(* Logix 5000 project; controller CIP_14485201 vendor 1 type 14 code 216 rev 38.11; software revision 38.01; part 2 of 12 *)

        [3].Setpoint[7] := 53.0, [3].Setpoint[8] := 63.0, [3].Setpoint[9] := 57.0, [3].Setpoint[10] := 43.0, [3].Setpoint[11] := 63.0, [3].Setpoint[13] := 85.0, [3].Setpoint[14] := 300.0, [3].Setpoint[15] := 900.0, [3].Setpoint[17] := 15.0, [3].Setpoint[18] := 14.0, [3].Setpoint[19] := 15.0, [3].Setpoint[20] := 45.0, [3].Setpoint[21] := 5.0, [3].Setpoint[22] := 15.0, [3].Setpoint[23] := 300.0, [3].Setpoint[25] := 10.0, [3].Setpoint[26] := 9.0, [3].Setpoint[27] := 10.0, [3].Setpoint[28] := 50.0, [3].Setpoint[29] := 3.0, [3].Setpoint[30] := 17.0, [3].Setpoint[31] := 300.0, [3].Setpoint[33] := 2.0, [3].Setpoint[34] := 900.0, [3].Setpoint[37] := 35.0, [3].Setpoint[41] := 5.0, [3].Setpoint[42] := 50.0, [3].Setpoint[43] := 5.0, [3].Setpoint[44] := 60.0, [3].Setpoint[45] := 50.0, [3].Setpoint[47] := 15.0, [3].Setpoint[49] := 180.0, [3].Setpoint[50] := 180.0, [3].Setpoint[52] := 30.0, [3].Setpoint[53] := 5.0, [3].Setpoint[54] := 5.0, [3].Setpoint[55] := 3.0, [3].Setpoint[57] := 300.0, [3].Name := 'RECIPE #3', [4].Setpoint[1] := 55.0, [4].Setpoint[2] := 65.0, [4].Setpoint[3] := 60.0, [4].Setpoint[4] := 45.0, [4].Setpoint[5] := 65.0, [4].Setpoint[7] := 53.0, [4].Setpoint[8] := 63.0, [4].Setpoint[9] := 57.0, [4].Setpoint[10] := 43.0, [4].Setpoint[11] := 63.0, [4].Setpoint[13] := 85.0, [4].Setpoint[14] := 300.0, [4].Setpoint[15] := 900.0, [4].Setpoint[17] := 15.0, [4].Setpoint[18] := 14.0, [4].Setpoint[19] := 15.0, [4].Setpoint[20] := 45.0, [4].Setpoint[21] := 5.0, [4].Setpoint[22] := 15.0, [4].Setpoint[23] := 300.0, [4].Setpoint[25] := 10.0,
        [4].Setpoint[26] := 9.0, [4].Setpoint[27] := 10.0, [4].Setpoint[28] := 50.0, [4].Setpoint[29] := 3.0, [4].Setpoint[30] := 17.0, [4].Setpoint[31] := 300.0, [4].Setpoint[33] := 2.0, [4].Setpoint[34] := 900.0, [4].Setpoint[37] := 35.0, [4].Setpoint[41] := 5.0, [4].Setpoint[42] := 50.0, [4].Setpoint[43] := 5.0, [4].Setpoint[44] := 60.0, [4].Setpoint[45] := 50.0, [4].Setpoint[47] := 15.0, [4].Setpoint[49] := 180.0, [4].Setpoint[50] := 180.0, [4].Setpoint[52] := 30.0, [4].Setpoint[53] := 5.0, [4].Setpoint[54] := 5.0, [4].Setpoint[55] := 3.0, [4].Setpoint[57] := 300.0, [4].Name := 'RECIPE #4', [5].Setpoint[1] := 55.0, [5].Setpoint[2] := 65.0, [5].Setpoint[3] := 60.0, [5].Setpoint[4] := 45.0, [5].Setpoint[5] := 65.0, [5].Setpoint[7] := 53.0, [5].Setpoint[8] := 63.0, [5].Setpoint[9] := 57.0, [5].Setpoint[10] := 43.0, [5].Setpoint[11] := 63.0, [5].Setpoint[13] := 85.0, [5].Setpoint[14] := 300.0, [5].Setpoint[15] := 900.0, [5].Setpoint[17] := 15.0, [5].Setpoint[18] := 14.0, [5].Setpoint[19] := 15.0, [5].Setpoint[20] := 45.0, [5].Setpoint[21] := 5.0, [5].Setpoint[22] := 15.0, [5].Setpoint[23] := 300.0, [5].Setpoint[25] := 10.0, [5].Setpoint[26] := 9.0, [5].Setpoint[27] := 10.0, [5].Setpoint[28] := 50.0, [5].Setpoint[29] := 3.0, [5].Setpoint[30] := 17.0, [5].Setpoint[31] := 300.0, [5].Setpoint[33] := 2.0, [5].Setpoint[34] := 900.0, [5].Setpoint[37] := 35.0, [5].Setpoint[41] := 5.0, [5].Setpoint[42] := 50.0, [5].Setpoint[43] := 5.0, [5].Setpoint[44] := 60.0, [5].Setpoint[45] := 50.0, [5].Setpoint[47] := 15.0, [5].Setpoint[49] := 180.0,
        [5].Setpoint[50] := 180.0, [5].Setpoint[52] := 30.0, [5].Setpoint[53] := 5.0, [5].Setpoint[54] := 5.0, [5].Setpoint[55] := 3.0, [5].Setpoint[57] := 300.0, [5].Name := 'RECIPE #5', [6].Setpoint[1] := 55.0, [6].Setpoint[2] := 65.0, [6].Setpoint[3] := 60.0, [6].Setpoint[4] := 45.0, [6].Setpoint[5] := 65.0, [6].Setpoint[7] := 53.0, [6].Setpoint[8] := 63.0, [6].Setpoint[9] := 57.0, [6].Setpoint[10] := 43.0, [6].Setpoint[11] := 63.0, [6].Setpoint[13] := 85.0, [6].Setpoint[14] := 300.0, [6].Setpoint[15] := 900.0, [6].Setpoint[17] := 15.0, [6].Setpoint[18] := 14.0, [6].Setpoint[19] := 15.0, [6].Setpoint[20] := 45.0, [6].Setpoint[21] := 5.0, [6].Setpoint[22] := 15.0, [6].Setpoint[23] := 300.0, [6].Setpoint[25] := 10.0, [6].Setpoint[26] := 9.0, [6].Setpoint[27] := 10.0, [6].Setpoint[28] := 50.0, [6].Setpoint[29] := 3.0, [6].Setpoint[30] := 17.0, [6].Setpoint[31] := 300.0, [6].Setpoint[33] := 2.0, [6].Setpoint[34] := 900.0, [6].Setpoint[37] := 35.0, [6].Setpoint[41] := 5.0, [6].Setpoint[42] := 50.0, [6].Setpoint[43] := 5.0, [6].Setpoint[44] := 60.0, [6].Setpoint[45] := 50.0, [6].Setpoint[47] := 15.0, [6].Setpoint[49] := 180.0, [6].Setpoint[50] := 180.0, [6].Setpoint[52] := 30.0, [6].Setpoint[53] := 5.0, [6].Setpoint[54] := 5.0, [6].Setpoint[55] := 3.0, [6].Setpoint[57] := 300.0, [6].Name := 'RECIPE #6', [7].Setpoint[1] := 55.0, [7].Setpoint[2] := 65.0, [7].Setpoint[3] := 60.0, [7].Setpoint[4] := 45.0, [7].Setpoint[5] := 65.0, [7].Setpoint[7] := 53.0, [7].Setpoint[8] := 63.0, [7].Setpoint[9] := 57.0, [7].Setpoint[10] := 43.0,
        [7].Setpoint[11] := 63.0, [7].Setpoint[13] := 85.0, [7].Setpoint[14] := 300.0, [7].Setpoint[15] := 900.0, [7].Setpoint[17] := 15.0, [7].Setpoint[18] := 14.0, [7].Setpoint[19] := 15.0, [7].Setpoint[20] := 45.0, [7].Setpoint[21] := 5.0, [7].Setpoint[22] := 15.0, [7].Setpoint[23] := 300.0, [7].Setpoint[25] := 10.0, [7].Setpoint[26] := 9.0, [7].Setpoint[27] := 10.0, [7].Setpoint[28] := 50.0, [7].Setpoint[29] := 3.0, [7].Setpoint[30] := 17.0, [7].Setpoint[31] := 300.0, [7].Setpoint[33] := 2.0, [7].Setpoint[34] := 900.0, [7].Setpoint[37] := 35.0, [7].Setpoint[41] := 5.0, [7].Setpoint[42] := 50.0, [7].Setpoint[43] := 5.0, [7].Setpoint[44] := 60.0, [7].Setpoint[45] := 50.0, [7].Setpoint[47] := 15.0, [7].Setpoint[49] := 180.0, [7].Setpoint[50] := 180.0, [7].Setpoint[52] := 30.0, [7].Setpoint[53] := 5.0, [7].Setpoint[54] := 5.0, [7].Setpoint[55] := 3.0, [7].Setpoint[57] := 300.0, [7].Name := 'RECIPE #7', [8].Setpoint[1] := 55.0, [8].Setpoint[2] := 65.0, [8].Setpoint[3] := 60.0, [8].Setpoint[4] := 45.0, [8].Setpoint[5] := 65.0, [8].Setpoint[7] := 53.0, [8].Setpoint[8] := 63.0, [8].Setpoint[9] := 57.0, [8].Setpoint[10] := 43.0, [8].Setpoint[11] := 63.0, [8].Setpoint[13] := 85.0, [8].Setpoint[14] := 300.0, [8].Setpoint[15] := 900.0, [8].Setpoint[17] := 15.0, [8].Setpoint[18] := 14.0, [8].Setpoint[19] := 15.0, [8].Setpoint[20] := 45.0, [8].Setpoint[21] := 5.0, [8].Setpoint[22] := 15.0, [8].Setpoint[23] := 300.0, [8].Setpoint[25] := 10.0, [8].Setpoint[26] := 9.0, [8].Setpoint[27] := 10.0, [8].Setpoint[28] := 50.0, [8].Setpoint[29] := 3.0,
        [8].Setpoint[30] := 17.0, [8].Setpoint[31] := 300.0, [8].Setpoint[33] := 2.0, [8].Setpoint[34] := 900.0, [8].Setpoint[37] := 35.0, [8].Setpoint[41] := 5.0, [8].Setpoint[42] := 50.0, [8].Setpoint[43] := 5.0, [8].Setpoint[44] := 60.0, [8].Setpoint[45] := 50.0, [8].Setpoint[47] := 15.0, [8].Setpoint[49] := 180.0, [8].Setpoint[50] := 180.0, [8].Setpoint[52] := 30.0, [8].Setpoint[53] := 5.0, [8].Setpoint[54] := 5.0, [8].Setpoint[55] := 3.0, [8].Setpoint[57] := 300.0, [8].Name := 'RECIPE #8', [9].Setpoint[1] := 55.0, [9].Setpoint[2] := 65.0, [9].Setpoint[3] := 60.0, [9].Setpoint[4] := 45.0, [9].Setpoint[5] := 65.0, [9].Setpoint[7] := 53.0, [9].Setpoint[8] := 63.0, [9].Setpoint[9] := 57.0, [9].Setpoint[10] := 43.0, [9].Setpoint[11] := 63.0, [9].Setpoint[13] := 85.0, [9].Setpoint[14] := 300.0, [9].Setpoint[15] := 900.0, [9].Setpoint[17] := 15.0, [9].Setpoint[18] := 14.0, [9].Setpoint[19] := 15.0, [9].Setpoint[20] := 45.0, [9].Setpoint[21] := 5.0, [9].Setpoint[22] := 15.0, [9].Setpoint[23] := 300.0, [9].Setpoint[25] := 10.0, [9].Setpoint[26] := 9.0, [9].Setpoint[27] := 10.0, [9].Setpoint[28] := 50.0, [9].Setpoint[29] := 3.0, [9].Setpoint[30] := 17.0, [9].Setpoint[31] := 300.0, [9].Setpoint[33] := 2.0, [9].Setpoint[34] := 900.0, [9].Setpoint[37] := 35.0, [9].Setpoint[41] := 5.0, [9].Setpoint[42] := 50.0, [9].Setpoint[43] := 5.0, [9].Setpoint[44] := 60.0, [9].Setpoint[45] := 50.0, [9].Setpoint[47] := 15.0, [9].Setpoint[49] := 180.0, [9].Setpoint[50] := 180.0, [9].Setpoint[52] := 30.0, [9].Setpoint[53] := 5.0, [9].Setpoint[54] := 5.0,
        [9].Setpoint[55] := 3.0, [9].Setpoint[57] := 300.0, [9].Name := 'RECIPE #9', [10].Setpoint[1] := 55.0, [10].Setpoint[2] := 65.0, [10].Setpoint[3] := 60.0, [10].Setpoint[4] := 45.0, [10].Setpoint[5] := 65.0, [10].Setpoint[7] := 53.0, [10].Setpoint[8] := 63.0, [10].Setpoint[9] := 57.0, [10].Setpoint[10] := 43.0, [10].Setpoint[11] := 63.0, [10].Setpoint[13] := 85.0, [10].Setpoint[14] := 300.0, [10].Setpoint[15] := 900.0, [10].Setpoint[17] := 15.0, [10].Setpoint[18] := 14.0, [10].Setpoint[19] := 15.0, [10].Setpoint[20] := 45.0, [10].Setpoint[21] := 5.0, [10].Setpoint[22] := 15.0, [10].Setpoint[23] := 300.0, [10].Setpoint[25] := 10.0, [10].Setpoint[26] := 9.0, [10].Setpoint[27] := 10.0, [10].Setpoint[28] := 50.0, [10].Setpoint[29] := 3.0, [10].Setpoint[30] := 17.0, [10].Setpoint[31] := 300.0, [10].Setpoint[33] := 2.0, [10].Setpoint[34] := 900.0, [10].Setpoint[37] := 35.0, [10].Setpoint[41] := 5.0, [10].Setpoint[42] := 50.0, [10].Setpoint[43] := 5.0, [10].Setpoint[44] := 60.0, [10].Setpoint[45] := 50.0, [10].Setpoint[47] := 15.0, [10].Setpoint[49] := 180.0, [10].Setpoint[50] := 180.0, [10].Setpoint[52] := 30.0, [10].Setpoint[53] := 5.0, [10].Setpoint[54] := 5.0, [10].Setpoint[55] := 3.0, [10].Setpoint[57] := 300.0, [10].Name := 'RECIPE #10', [11].Setpoint[1] := 55.0, [11].Setpoint[2] := 65.0, [11].Setpoint[3] := 60.0, [11].Setpoint[4] := 45.0, [11].Setpoint[5] := 65.0, [11].Setpoint[7] := 53.0, [11].Setpoint[8] := 63.0, [11].Setpoint[9] := 57.0, [11].Setpoint[10] := 43.0, [11].Setpoint[11] := 63.0, [11].Setpoint[13] := 85.0, [11].Setpoint[14] := 300.0, [11].Setpoint[15] := 900.0,
        [11].Setpoint[17] := 15.0, [11].Setpoint[18] := 14.0, [11].Setpoint[19] := 15.0, [11].Setpoint[20] := 45.0, [11].Setpoint[21] := 5.0, [11].Setpoint[22] := 15.0, [11].Setpoint[23] := 300.0, [11].Setpoint[25] := 10.0, [11].Setpoint[26] := 9.0, [11].Setpoint[27] := 10.0, [11].Setpoint[28] := 50.0, [11].Setpoint[29] := 3.0, [11].Setpoint[30] := 17.0, [11].Setpoint[31] := 300.0, [11].Setpoint[33] := 2.0, [11].Setpoint[34] := 900.0, [11].Setpoint[37] := 35.0, [11].Setpoint[41] := 5.0, [11].Setpoint[42] := 50.0, [11].Setpoint[43] := 5.0, [11].Setpoint[44] := 60.0, [11].Setpoint[45] := 50.0, [11].Setpoint[47] := 15.0, [11].Setpoint[49] := 180.0, [11].Setpoint[50] := 180.0, [11].Setpoint[52] := 30.0, [11].Setpoint[53] := 5.0, [11].Setpoint[54] := 5.0, [11].Setpoint[55] := 3.0, [11].Setpoint[57] := 300.0, [11].Name := 'RECIPE #11', [12].Setpoint[1] := 55.0, [12].Setpoint[2] := 65.0, [12].Setpoint[3] := 60.0, [12].Setpoint[4] := 45.0, [12].Setpoint[5] := 65.0, [12].Setpoint[7] := 53.0, [12].Setpoint[8] := 63.0, [12].Setpoint[9] := 57.0, [12].Setpoint[10] := 43.0, [12].Setpoint[11] := 63.0, [12].Setpoint[13] := 85.0, [12].Setpoint[14] := 300.0, [12].Setpoint[15] := 900.0, [12].Setpoint[17] := 15.0, [12].Setpoint[18] := 14.0, [12].Setpoint[19] := 15.0, [12].Setpoint[20] := 45.0, [12].Setpoint[21] := 5.0, [12].Setpoint[22] := 15.0, [12].Setpoint[23] := 300.0, [12].Setpoint[25] := 10.0, [12].Setpoint[26] := 9.0, [12].Setpoint[27] := 10.0, [12].Setpoint[28] := 50.0, [12].Setpoint[29] := 3.0, [12].Setpoint[30] := 17.0, [12].Setpoint[31] := 300.0, [12].Setpoint[33] := 2.0, [12].Setpoint[34] := 900.0,
        [12].Setpoint[37] := 35.0, [12].Setpoint[41] := 5.0, [12].Setpoint[42] := 50.0, [12].Setpoint[43] := 5.0, [12].Setpoint[44] := 60.0, [12].Setpoint[45] := 50.0, [12].Setpoint[47] := 15.0, [12].Setpoint[49] := 180.0, [12].Setpoint[50] := 180.0, [12].Setpoint[52] := 30.0, [12].Setpoint[53] := 5.0, [12].Setpoint[54] := 5.0, [12].Setpoint[55] := 3.0, [12].Setpoint[57] := 300.0, [12].Name := 'RECIPE #12', [13].Setpoint[1] := 55.0, [13].Setpoint[2] := 65.0, [13].Setpoint[3] := 60.0, [13].Setpoint[4] := 45.0, [13].Setpoint[5] := 65.0, [13].Setpoint[7] := 53.0, [13].Setpoint[8] := 63.0, [13].Setpoint[9] := 57.0, [13].Setpoint[10] := 43.0, [13].Setpoint[11] := 63.0, [13].Setpoint[13] := 85.0, [13].Setpoint[14] := 300.0, [13].Setpoint[15] := 900.0, [13].Setpoint[17] := 15.0, [13].Setpoint[18] := 14.0, [13].Setpoint[19] := 15.0, [13].Setpoint[20] := 45.0, [13].Setpoint[21] := 5.0, [13].Setpoint[22] := 15.0, [13].Setpoint[23] := 300.0, [13].Setpoint[25] := 10.0, [13].Setpoint[26] := 9.0, [13].Setpoint[27] := 10.0, [13].Setpoint[28] := 50.0, [13].Setpoint[29] := 3.0, [13].Setpoint[30] := 17.0, [13].Setpoint[31] := 300.0, [13].Setpoint[33] := 2.0, [13].Setpoint[34] := 900.0, [13].Setpoint[37] := 35.0, [13].Setpoint[41] := 5.0, [13].Setpoint[42] := 50.0, [13].Setpoint[43] := 5.0, [13].Setpoint[44] := 60.0, [13].Setpoint[45] := 50.0, [13].Setpoint[47] := 15.0, [13].Setpoint[49] := 180.0, [13].Setpoint[50] := 180.0, [13].Setpoint[52] := 30.0, [13].Setpoint[53] := 5.0, [13].Setpoint[54] := 5.0, [13].Setpoint[55] := 3.0, [13].Setpoint[57] := 300.0, [13].Name := 'RECIPE #13', [14].Setpoint[1] := 55.0,
        [14].Setpoint[2] := 65.0, [14].Setpoint[3] := 60.0, [14].Setpoint[4] := 45.0, [14].Setpoint[5] := 65.0, [14].Setpoint[7] := 53.0, [14].Setpoint[8] := 63.0, [14].Setpoint[9] := 57.0, [14].Setpoint[10] := 43.0, [14].Setpoint[11] := 63.0, [14].Setpoint[13] := 85.0, [14].Setpoint[14] := 300.0, [14].Setpoint[15] := 900.0, [14].Setpoint[17] := 15.0, [14].Setpoint[18] := 14.0, [14].Setpoint[19] := 15.0, [14].Setpoint[20] := 45.0, [14].Setpoint[21] := 5.0, [14].Setpoint[22] := 15.0, [14].Setpoint[23] := 300.0, [14].Setpoint[25] := 10.0, [14].Setpoint[26] := 9.0, [14].Setpoint[27] := 10.0, [14].Setpoint[28] := 50.0, [14].Setpoint[29] := 3.0, [14].Setpoint[30] := 17.0, [14].Setpoint[31] := 300.0, [14].Setpoint[33] := 2.0, [14].Setpoint[34] := 900.0, [14].Setpoint[37] := 35.0, [14].Setpoint[41] := 5.0, [14].Setpoint[42] := 50.0, [14].Setpoint[43] := 5.0, [14].Setpoint[44] := 60.0, [14].Setpoint[45] := 50.0, [14].Setpoint[47] := 15.0, [14].Setpoint[49] := 180.0, [14].Setpoint[50] := 180.0, [14].Setpoint[52] := 30.0, [14].Setpoint[53] := 5.0, [14].Setpoint[54] := 5.0, [14].Setpoint[55] := 3.0, [14].Setpoint[57] := 300.0, [14].Name := 'RECIPE #14', [15].Setpoint[1] := 55.0, [15].Setpoint[2] := 65.0, [15].Setpoint[3] := 60.0, [15].Setpoint[4] := 45.0, [15].Setpoint[5] := 65.0, [15].Setpoint[7] := 53.0, [15].Setpoint[8] := 63.0, [15].Setpoint[9] := 57.0, [15].Setpoint[10] := 43.0, [15].Setpoint[11] := 63.0, [15].Setpoint[13] := 85.0, [15].Setpoint[14] := 300.0, [15].Setpoint[15] := 900.0, [15].Setpoint[17] := 15.0, [15].Setpoint[18] := 14.0, [15].Setpoint[19] := 15.0, [15].Setpoint[20] := 45.0,
        [15].Setpoint[21] := 5.0, [15].Setpoint[22] := 15.0, [15].Setpoint[23] := 300.0, [15].Setpoint[25] := 10.0, [15].Setpoint[26] := 9.0, [15].Setpoint[27] := 10.0, [15].Setpoint[28] := 50.0, [15].Setpoint[29] := 3.0, [15].Setpoint[30] := 17.0, [15].Setpoint[31] := 300.0, [15].Setpoint[33] := 2.0, [15].Setpoint[34] := 900.0, [15].Setpoint[37] := 35.0, [15].Setpoint[41] := 5.0, [15].Setpoint[42] := 50.0, [15].Setpoint[43] := 5.0, [15].Setpoint[44] := 60.0, [15].Setpoint[45] := 50.0, [15].Setpoint[47] := 15.0, [15].Setpoint[49] := 180.0, [15].Setpoint[50] := 180.0, [15].Setpoint[52] := 30.0, [15].Setpoint[53] := 5.0, [15].Setpoint[54] := 5.0, [15].Setpoint[55] := 3.0, [15].Setpoint[57] := 300.0, [15].Name := 'RECIPE #15', [16].Setpoint[1] := 55.0, [16].Setpoint[2] := 65.0, [16].Setpoint[3] := 60.0, [16].Setpoint[4] := 45.0, [16].Setpoint[5] := 65.0, [16].Setpoint[7] := 53.0, [16].Setpoint[8] := 63.0, [16].Setpoint[9] := 57.0, [16].Setpoint[10] := 43.0, [16].Setpoint[11] := 63.0, [16].Setpoint[13] := 85.0, [16].Setpoint[14] := 300.0, [16].Setpoint[15] := 900.0, [16].Setpoint[17] := 15.0, [16].Setpoint[18] := 14.0, [16].Setpoint[19] := 15.0, [16].Setpoint[20] := 45.0, [16].Setpoint[21] := 5.0, [16].Setpoint[22] := 15.0, [16].Setpoint[23] := 300.0, [16].Setpoint[25] := 10.0, [16].Setpoint[26] := 9.0, [16].Setpoint[27] := 10.0, [16].Setpoint[28] := 50.0, [16].Setpoint[29] := 3.0, [16].Setpoint[30] := 17.0, [16].Setpoint[31] := 300.0, [16].Setpoint[33] := 2.0, [16].Setpoint[34] := 900.0, [16].Setpoint[37] := 35.0, [16].Setpoint[41] := 5.0, [16].Setpoint[42] := 50.0, [16].Setpoint[43] := 5.0,
        [16].Setpoint[44] := 60.0, [16].Setpoint[45] := 50.0, [16].Setpoint[47] := 15.0, [16].Setpoint[49] := 180.0, [16].Setpoint[50] := 180.0, [16].Setpoint[52] := 30.0, [16].Setpoint[53] := 5.0, [16].Setpoint[54] := 5.0, [16].Setpoint[55] := 3.0, [16].Setpoint[57] := 300.0, [16].Name := 'RECIPE #16', [17].Setpoint[1] := 55.0, [17].Setpoint[2] := 65.0, [17].Setpoint[3] := 60.0, [17].Setpoint[4] := 45.0, [17].Setpoint[5] := 65.0, [17].Setpoint[7] := 53.0, [17].Setpoint[8] := 63.0, [17].Setpoint[9] := 57.0, [17].Setpoint[10] := 43.0, [17].Setpoint[11] := 63.0, [17].Setpoint[13] := 85.0, [17].Setpoint[14] := 300.0, [17].Setpoint[15] := 900.0, [17].Setpoint[17] := 15.0, [17].Setpoint[18] := 14.0, [17].Setpoint[19] := 15.0, [17].Setpoint[20] := 45.0, [17].Setpoint[21] := 5.0, [17].Setpoint[22] := 15.0, [17].Setpoint[23] := 300.0, [17].Setpoint[25] := 10.0, [17].Setpoint[26] := 9.0, [17].Setpoint[27] := 10.0, [17].Setpoint[28] := 50.0, [17].Setpoint[29] := 3.0, [17].Setpoint[30] := 17.0, [17].Setpoint[31] := 300.0, [17].Setpoint[33] := 2.0, [17].Setpoint[34] := 900.0, [17].Setpoint[37] := 35.0, [17].Setpoint[41] := 5.0, [17].Setpoint[42] := 50.0, [17].Setpoint[43] := 5.0, [17].Setpoint[44] := 60.0, [17].Setpoint[45] := 50.0, [17].Setpoint[47] := 15.0, [17].Setpoint[49] := 180.0, [17].Setpoint[50] := 180.0, [17].Setpoint[52] := 30.0, [17].Setpoint[53] := 5.0, [17].Setpoint[54] := 5.0, [17].Setpoint[55] := 3.0, [17].Setpoint[57] := 300.0, [17].Name := 'RECIPE #17', [18].Setpoint[1] := 55.0, [18].Setpoint[2] := 65.0, [18].Setpoint[3] := 60.0, [18].Setpoint[4] := 45.0, [18].Setpoint[5] := 65.0,
        [18].Setpoint[7] := 53.0, [18].Setpoint[8] := 63.0, [18].Setpoint[9] := 57.0, [18].Setpoint[10] := 43.0, [18].Setpoint[11] := 63.0, [18].Setpoint[13] := 85.0, [18].Setpoint[14] := 300.0, [18].Setpoint[15] := 900.0, [18].Setpoint[17] := 15.0, [18].Setpoint[18] := 14.0, [18].Setpoint[19] := 15.0, [18].Setpoint[20] := 45.0, [18].Setpoint[21] := 5.0, [18].Setpoint[22] := 15.0, [18].Setpoint[23] := 300.0, [18].Setpoint[25] := 10.0, [18].Setpoint[26] := 9.0, [18].Setpoint[27] := 10.0, [18].Setpoint[28] := 50.0, [18].Setpoint[29] := 3.0, [18].Setpoint[30] := 17.0, [18].Setpoint[31] := 300.0, [18].Setpoint[33] := 2.0, [18].Setpoint[34] := 900.0, [18].Setpoint[37] := 35.0, [18].Setpoint[41] := 5.0, [18].Setpoint[42] := 50.0, [18].Setpoint[43] := 5.0, [18].Setpoint[44] := 60.0, [18].Setpoint[45] := 50.0, [18].Setpoint[47] := 15.0, [18].Setpoint[49] := 180.0, [18].Setpoint[50] := 180.0, [18].Setpoint[52] := 30.0, [18].Setpoint[53] := 5.0, [18].Setpoint[54] := 5.0, [18].Setpoint[55] := 3.0, [18].Setpoint[57] := 300.0, [18].Name := 'RECIPE #18', [19].Setpoint[1] := 55.0, [19].Setpoint[2] := 65.0, [19].Setpoint[3] := 60.0, [19].Setpoint[4] := 45.0, [19].Setpoint[5] := 65.0, [19].Setpoint[7] := 53.0, [19].Setpoint[8] := 63.0, [19].Setpoint[9] := 57.0, [19].Setpoint[10] := 43.0, [19].Setpoint[11] := 63.0, [19].Setpoint[13] := 85.0, [19].Setpoint[14] := 300.0, [19].Setpoint[15] := 900.0, [19].Setpoint[17] := 15.0, [19].Setpoint[18] := 14.0, [19].Setpoint[19] := 15.0, [19].Setpoint[20] := 45.0, [19].Setpoint[21] := 5.0, [19].Setpoint[22] := 15.0, [19].Setpoint[23] := 300.0, [19].Setpoint[25] := 10.0,
        [19].Setpoint[26] := 9.0, [19].Setpoint[27] := 10.0, [19].Setpoint[28] := 50.0, [19].Setpoint[29] := 3.0, [19].Setpoint[30] := 17.0, [19].Setpoint[31] := 300.0, [19].Setpoint[33] := 2.0, [19].Setpoint[34] := 900.0, [19].Setpoint[37] := 35.0, [19].Setpoint[41] := 5.0, [19].Setpoint[42] := 50.0, [19].Setpoint[43] := 5.0, [19].Setpoint[44] := 60.0, [19].Setpoint[45] := 50.0, [19].Setpoint[47] := 15.0, [19].Setpoint[49] := 180.0, [19].Setpoint[50] := 180.0, [19].Setpoint[52] := 30.0, [19].Setpoint[53] := 5.0, [19].Setpoint[54] := 5.0, [19].Setpoint[55] := 3.0, [19].Setpoint[57] := 300.0, [19].Name := 'RECIPE #19', [20].Setpoint[1] := 55.0, [20].Setpoint[2] := 65.0, [20].Setpoint[3] := 60.0, [20].Setpoint[4] := 45.0, [20].Setpoint[5] := 65.0, [20].Setpoint[7] := 53.0, [20].Setpoint[8] := 63.0, [20].Setpoint[9] := 57.0, [20].Setpoint[10] := 43.0, [20].Setpoint[11] := 63.0, [20].Setpoint[13] := 85.0, [20].Setpoint[14] := 300.0, [20].Setpoint[15] := 900.0, [20].Setpoint[17] := 15.0, [20].Setpoint[18] := 14.0, [20].Setpoint[19] := 15.0, [20].Setpoint[20] := 45.0, [20].Setpoint[21] := 5.0, [20].Setpoint[22] := 15.0, [20].Setpoint[23] := 300.0, [20].Setpoint[25] := 10.0, [20].Setpoint[26] := 9.0, [20].Setpoint[27] := 10.0, [20].Setpoint[28] := 50.0, [20].Setpoint[29] := 3.0, [20].Setpoint[30] := 17.0, [20].Setpoint[31] := 300.0, [20].Setpoint[33] := 2.0, [20].Setpoint[34] := 900.0, [20].Setpoint[37] := 35.0, [20].Setpoint[41] := 5.0, [20].Setpoint[42] := 50.0, [20].Setpoint[43] := 5.0, [20].Setpoint[44] := 60.0, [20].Setpoint[45] := 50.0, [20].Setpoint[47] := 15.0, [20].Setpoint[49] := 180.0,
        [20].Setpoint[50] := 180.0, [20].Setpoint[52] := 30.0, [20].Setpoint[53] := 5.0, [20].Setpoint[54] := 5.0, [20].Setpoint[55] := 3.0, [20].Setpoint[57] := 300.0, [20].Name := 'RECIPE #20', [21].Setpoint[1] := 55.0, [21].Setpoint[2] := 65.0, [21].Setpoint[3] := 60.0, [21].Setpoint[4] := 45.0, [21].Setpoint[5] := 65.0, [21].Setpoint[7] := 53.0, [21].Setpoint[8] := 63.0, [21].Setpoint[9] := 57.0, [21].Setpoint[10] := 43.0, [21].Setpoint[11] := 63.0, [21].Setpoint[13] := 85.0, [21].Setpoint[14] := 300.0, [21].Setpoint[15] := 900.0, [21].Setpoint[17] := 15.0, [21].Setpoint[18] := 14.0, [21].Setpoint[19] := 15.0, [21].Setpoint[20] := 45.0, [21].Setpoint[21] := 5.0, [21].Setpoint[22] := 15.0, [21].Setpoint[23] := 300.0, [21].Setpoint[25] := 10.0, [21].Setpoint[26] := 9.0, [21].Setpoint[27] := 10.0, [21].Setpoint[28] := 50.0, [21].Setpoint[29] := 3.0, [21].Setpoint[30] := 17.0, [21].Setpoint[31] := 300.0, [21].Setpoint[33] := 2.0, [21].Setpoint[34] := 900.0, [21].Setpoint[37] := 35.0, [21].Setpoint[41] := 5.0, [21].Setpoint[42] := 50.0, [21].Setpoint[43] := 5.0, [21].Setpoint[44] := 60.0, [21].Setpoint[45] := 50.0, [21].Setpoint[47] := 15.0, [21].Setpoint[49] := 180.0, [21].Setpoint[50] := 180.0, [21].Setpoint[52] := 30.0, [21].Setpoint[53] := 5.0, [21].Setpoint[54] := 5.0, [21].Setpoint[55] := 3.0, [21].Setpoint[57] := 300.0, [21].Name := 'RECIPE #21', [22].Setpoint[1] := 55.0, [22].Setpoint[2] := 65.0, [22].Setpoint[3] := 60.0, [22].Setpoint[4] := 45.0, [22].Setpoint[5] := 65.0, [22].Setpoint[7] := 53.0, [22].Setpoint[8] := 63.0, [22].Setpoint[9] := 57.0, [22].Setpoint[10] := 43.0,
        [22].Setpoint[11] := 63.0, [22].Setpoint[13] := 85.0, [22].Setpoint[14] := 300.0, [22].Setpoint[15] := 900.0, [22].Setpoint[17] := 15.0, [22].Setpoint[18] := 14.0, [22].Setpoint[19] := 15.0, [22].Setpoint[20] := 45.0, [22].Setpoint[21] := 5.0, [22].Setpoint[22] := 15.0, [22].Setpoint[23] := 300.0, [22].Setpoint[25] := 10.0, [22].Setpoint[26] := 9.0, [22].Setpoint[27] := 10.0, [22].Setpoint[28] := 50.0, [22].Setpoint[29] := 3.0, [22].Setpoint[30] := 17.0, [22].Setpoint[31] := 300.0, [22].Setpoint[33] := 2.0, [22].Setpoint[34] := 900.0, [22].Setpoint[37] := 35.0, [22].Setpoint[41] := 5.0, [22].Setpoint[42] := 50.0, [22].Setpoint[43] := 5.0, [22].Setpoint[44] := 60.0, [22].Setpoint[45] := 50.0, [22].Setpoint[47] := 15.0, [22].Setpoint[49] := 180.0, [22].Setpoint[50] := 180.0, [22].Setpoint[52] := 30.0, [22].Setpoint[53] := 5.0, [22].Setpoint[54] := 5.0, [22].Setpoint[55] := 3.0, [22].Setpoint[57] := 300.0, [22].Name := 'RECIPE #22', [23].Setpoint[1] := 55.0, [23].Setpoint[2] := 65.0, [23].Setpoint[3] := 60.0, [23].Setpoint[4] := 45.0, [23].Setpoint[5] := 65.0, [23].Setpoint[7] := 53.0, [23].Setpoint[8] := 63.0, [23].Setpoint[9] := 57.0, [23].Setpoint[10] := 43.0, [23].Setpoint[11] := 63.0, [23].Setpoint[13] := 85.0, [23].Setpoint[14] := 300.0, [23].Setpoint[15] := 900.0, [23].Setpoint[17] := 15.0, [23].Setpoint[18] := 14.0, [23].Setpoint[19] := 15.0, [23].Setpoint[20] := 45.0, [23].Setpoint[21] := 5.0, [23].Setpoint[22] := 15.0, [23].Setpoint[23] := 300.0, [23].Setpoint[25] := 10.0, [23].Setpoint[26] := 9.0, [23].Setpoint[27] := 10.0, [23].Setpoint[28] := 50.0, [23].Setpoint[29] := 3.0,
        [23].Setpoint[30] := 17.0, [23].Setpoint[31] := 300.0, [23].Setpoint[33] := 2.0, [23].Setpoint[34] := 900.0, [23].Setpoint[37] := 35.0, [23].Setpoint[41] := 5.0, [23].Setpoint[42] := 50.0, [23].Setpoint[43] := 5.0, [23].Setpoint[44] := 60.0, [23].Setpoint[45] := 50.0, [23].Setpoint[47] := 15.0, [23].Setpoint[49] := 180.0, [23].Setpoint[50] := 180.0, [23].Setpoint[52] := 30.0, [23].Setpoint[53] := 5.0, [23].Setpoint[54] := 5.0, [23].Setpoint[55] := 3.0, [23].Setpoint[57] := 300.0, [23].Name := 'RECIPE #23', [24].OpCode[88] := 2, [24].Setpoint[1] := 55.0, [24].Setpoint[2] := 65.0, [24].Setpoint[3] := 60.0, [24].Setpoint[4] := 45.0, [24].Setpoint[5] := 65.0, [24].Setpoint[7] := 53.0, [24].Setpoint[8] := 63.0, [24].Setpoint[9] := 57.0, [24].Setpoint[10] := 43.0, [24].Setpoint[11] := 63.0, [24].Setpoint[13] := 85.0, [24].Setpoint[14] := 300.0, [24].Setpoint[15] := 900.0, [24].Setpoint[17] := 15.0, [24].Setpoint[18] := 14.0, [24].Setpoint[19] := 15.0, [24].Setpoint[20] := 45.0, [24].Setpoint[21] := 5.0, [24].Setpoint[22] := 15.0, [24].Setpoint[23] := 300.0, [24].Setpoint[25] := 10.0, [24].Setpoint[26] := 9.0, [24].Setpoint[27] := 10.0, [24].Setpoint[28] := 50.0, [24].Setpoint[29] := 3.0, [24].Setpoint[30] := 17.0, [24].Setpoint[31] := 300.0, [24].Setpoint[33] := 2.0, [24].Setpoint[34] := 900.0, [24].Setpoint[37] := 35.0, [24].Setpoint[41] := 5.0, [24].Setpoint[42] := 50.0, [24].Setpoint[43] := 5.0, [24].Setpoint[44] := 60.0, [24].Setpoint[45] := 50.0, [24].Setpoint[47] := 15.0, [24].Setpoint[49] := 180.0, [24].Setpoint[50] := 180.0, [24].Setpoint[52] := 30.0, [24].Setpoint[53] := 5.0,
        [24].Setpoint[54] := 5.0, [24].Setpoint[55] := 3.0, [24].Setpoint[57] := 300.0, [24].Name := 'RECIPE #24', [25].Setpoint[1] := 55.0, [25].Setpoint[2] := 65.0, [25].Setpoint[3] := 60.0, [25].Setpoint[4] := 45.0, [25].Setpoint[5] := 65.0, [25].Setpoint[7] := 53.0, [25].Setpoint[8] := 63.0, [25].Setpoint[9] := 57.0, [25].Setpoint[10] := 43.0, [25].Setpoint[11] := 63.0, [25].Setpoint[13] := 85.0, [25].Setpoint[14] := 300.0, [25].Setpoint[15] := 900.0, [25].Setpoint[17] := 15.0, [25].Setpoint[18] := 14.0, [25].Setpoint[19] := 15.0, [25].Setpoint[20] := 45.0, [25].Setpoint[21] := 5.0, [25].Setpoint[22] := 15.0, [25].Setpoint[23] := 300.0, [25].Setpoint[25] := 10.0, [25].Setpoint[26] := 9.0, [25].Setpoint[27] := 10.0, [25].Setpoint[28] := 50.0, [25].Setpoint[29] := 3.0, [25].Setpoint[30] := 17.0, [25].Setpoint[31] := 300.0, [25].Setpoint[33] := 2.0, [25].Setpoint[34] := 900.0, [25].Setpoint[37] := 35.0, [25].Setpoint[41] := 5.0, [25].Setpoint[42] := 50.0, [25].Setpoint[43] := 5.0, [25].Setpoint[44] := 60.0, [25].Setpoint[45] := 50.0, [25].Setpoint[47] := 15.0, [25].Setpoint[49] := 180.0, [25].Setpoint[50] := 180.0, [25].Setpoint[52] := 30.0, [25].Setpoint[53] := 5.0, [25].Setpoint[54] := 5.0, [25].Setpoint[55] := 3.0, [25].Setpoint[57] := 300.0, [25].Name := 'RECIPE #25', [26].Setpoint[1] := 55.0, [26].Setpoint[2] := 65.0, [26].Setpoint[3] := 60.0, [26].Setpoint[4] := 45.0, [26].Setpoint[5] := 65.0, [26].Setpoint[7] := 53.0, [26].Setpoint[8] := 63.0, [26].Setpoint[9] := 57.0, [26].Setpoint[10] := 43.0, [26].Setpoint[11] := 63.0, [26].Setpoint[13] := 85.0, [26].Setpoint[14] := 300.0,
        [26].Setpoint[15] := 900.0, [26].Setpoint[17] := 15.0, [26].Setpoint[18] := 14.0, [26].Setpoint[19] := 15.0, [26].Setpoint[20] := 45.0, [26].Setpoint[21] := 5.0, [26].Setpoint[22] := 15.0, [26].Setpoint[23] := 300.0, [26].Setpoint[25] := 10.0, [26].Setpoint[26] := 9.0, [26].Setpoint[27] := 10.0, [26].Setpoint[28] := 50.0, [26].Setpoint[29] := 3.0, [26].Setpoint[30] := 17.0, [26].Setpoint[31] := 300.0, [26].Setpoint[33] := 2.0, [26].Setpoint[34] := 900.0, [26].Setpoint[37] := 35.0, [26].Setpoint[41] := 5.0, [26].Setpoint[42] := 50.0, [26].Setpoint[43] := 5.0, [26].Setpoint[44] := 60.0, [26].Setpoint[45] := 50.0, [26].Setpoint[47] := 15.0, [26].Setpoint[49] := 180.0, [26].Setpoint[50] := 180.0, [26].Setpoint[52] := 30.0, [26].Setpoint[53] := 5.0, [26].Setpoint[54] := 5.0, [26].Setpoint[55] := 3.0, [26].Setpoint[57] := 300.0, [26].Name := 'RECIPE #26', [27].Setpoint[1] := 55.0, [27].Setpoint[2] := 65.0, [27].Setpoint[3] := 60.0, [27].Setpoint[4] := 45.0, [27].Setpoint[5] := 65.0, [27].Setpoint[7] := 53.0, [27].Setpoint[8] := 63.0, [27].Setpoint[9] := 57.0, [27].Setpoint[10] := 43.0, [27].Setpoint[11] := 63.0, [27].Setpoint[13] := 85.0, [27].Setpoint[14] := 300.0, [27].Setpoint[15] := 900.0, [27].Setpoint[17] := 15.0, [27].Setpoint[18] := 14.0, [27].Setpoint[19] := 15.0, [27].Setpoint[20] := 45.0, [27].Setpoint[21] := 5.0, [27].Setpoint[22] := 15.0, [27].Setpoint[23] := 300.0, [27].Setpoint[25] := 10.0, [27].Setpoint[26] := 9.0, [27].Setpoint[27] := 10.0, [27].Setpoint[28] := 50.0, [27].Setpoint[29] := 3.0, [27].Setpoint[30] := 17.0, [27].Setpoint[31] := 300.0, [27].Setpoint[33] := 2.0,
        [27].Setpoint[34] := 900.0, [27].Setpoint[37] := 35.0, [27].Setpoint[41] := 5.0, [27].Setpoint[42] := 50.0, [27].Setpoint[43] := 5.0, [27].Setpoint[44] := 60.0, [27].Setpoint[45] := 50.0, [27].Setpoint[47] := 15.0, [27].Setpoint[49] := 180.0, [27].Setpoint[50] := 180.0, [27].Setpoint[52] := 30.0, [27].Setpoint[53] := 5.0, [27].Setpoint[54] := 5.0, [27].Setpoint[55] := 3.0, [27].Setpoint[57] := 300.0, [27].Name := 'RECIPE #27', [28].Setpoint[1] := 55.0, [28].Setpoint[2] := 65.0, [28].Setpoint[3] := 60.0, [28].Setpoint[4] := 45.0, [28].Setpoint[5] := 65.0, [28].Setpoint[7] := 53.0, [28].Setpoint[8] := 63.0, [28].Setpoint[9] := 57.0, [28].Setpoint[10] := 43.0, [28].Setpoint[11] := 63.0, [28].Setpoint[13] := 85.0, [28].Setpoint[14] := 300.0, [28].Setpoint[15] := 900.0, [28].Setpoint[17] := 15.0, [28].Setpoint[18] := 14.0, [28].Setpoint[19] := 15.0, [28].Setpoint[20] := 45.0, [28].Setpoint[21] := 5.0, [28].Setpoint[22] := 15.0, [28].Setpoint[23] := 300.0, [28].Setpoint[25] := 10.0, [28].Setpoint[26] := 9.0, [28].Setpoint[27] := 10.0, [28].Setpoint[28] := 50.0, [28].Setpoint[29] := 3.0, [28].Setpoint[30] := 17.0, [28].Setpoint[31] := 300.0, [28].Setpoint[33] := 2.0, [28].Setpoint[34] := 900.0, [28].Setpoint[37] := 35.0, [28].Setpoint[41] := 5.0, [28].Setpoint[42] := 50.0, [28].Setpoint[43] := 5.0, [28].Setpoint[44] := 60.0, [28].Setpoint[45] := 50.0, [28].Setpoint[47] := 15.0, [28].Setpoint[49] := 180.0, [28].Setpoint[50] := 180.0, [28].Setpoint[52] := 30.0, [28].Setpoint[53] := 5.0, [28].Setpoint[54] := 5.0, [28].Setpoint[55] := 3.0, [28].Setpoint[57] := 300.0, [28].Name := 'RECIPE #28',
        [29].Setpoint[1] := 55.0, [29].Setpoint[2] := 65.0, [29].Setpoint[3] := 60.0, [29].Setpoint[4] := 45.0, [29].Setpoint[5] := 65.0, [29].Setpoint[7] := 53.0, [29].Setpoint[8] := 63.0, [29].Setpoint[9] := 57.0, [29].Setpoint[10] := 43.0, [29].Setpoint[11] := 63.0, [29].Setpoint[13] := 85.0, [29].Setpoint[14] := 300.0, [29].Setpoint[15] := 900.0, [29].Setpoint[17] := 15.0, [29].Setpoint[18] := 14.0, [29].Setpoint[19] := 15.0, [29].Setpoint[20] := 45.0, [29].Setpoint[21] := 5.0, [29].Setpoint[22] := 15.0, [29].Setpoint[23] := 300.0, [29].Setpoint[25] := 10.0, [29].Setpoint[26] := 9.0, [29].Setpoint[27] := 10.0, [29].Setpoint[28] := 50.0, [29].Setpoint[29] := 3.0, [29].Setpoint[30] := 17.0, [29].Setpoint[31] := 300.0, [29].Setpoint[33] := 2.0, [29].Setpoint[34] := 900.0, [29].Setpoint[37] := 35.0, [29].Setpoint[41] := 5.0, [29].Setpoint[42] := 50.0, [29].Setpoint[43] := 5.0, [29].Setpoint[44] := 60.0, [29].Setpoint[45] := 50.0, [29].Setpoint[47] := 15.0, [29].Setpoint[49] := 180.0, [29].Setpoint[50] := 180.0, [29].Setpoint[52] := 30.0, [29].Setpoint[53] := 5.0, [29].Setpoint[54] := 5.0, [29].Setpoint[55] := 3.0, [29].Setpoint[57] := 300.0, [29].Name := 'RECIPE #29', [30].Setpoint[1] := 55.0, [30].Setpoint[2] := 65.0, [30].Setpoint[3] := 60.0, [30].Setpoint[4] := 45.0, [30].Setpoint[5] := 65.0, [30].Setpoint[7] := 53.0, [30].Setpoint[8] := 63.0, [30].Setpoint[9] := 57.0, [30].Setpoint[10] := 43.0, [30].Setpoint[11] := 63.0, [30].Setpoint[13] := 85.0, [30].Setpoint[14] := 300.0, [30].Setpoint[15] := 900.0, [30].Setpoint[17] := 15.0, [30].Setpoint[18] := 14.0, [30].Setpoint[19] := 15.0,
        [30].Setpoint[20] := 45.0, [30].Setpoint[21] := 5.0, [30].Setpoint[22] := 15.0, [30].Setpoint[23] := 300.0, [30].Setpoint[25] := 10.0, [30].Setpoint[26] := 9.0, [30].Setpoint[27] := 10.0, [30].Setpoint[28] := 50.0, [30].Setpoint[29] := 3.0, [30].Setpoint[30] := 17.0, [30].Setpoint[31] := 300.0, [30].Setpoint[33] := 2.0, [30].Setpoint[34] := 900.0, [30].Setpoint[37] := 35.0, [30].Setpoint[41] := 5.0, [30].Setpoint[42] := 50.0, [30].Setpoint[43] := 5.0, [30].Setpoint[44] := 60.0, [30].Setpoint[45] := 50.0, [30].Setpoint[47] := 15.0, [30].Setpoint[49] := 180.0, [30].Setpoint[50] := 180.0, [30].Setpoint[52] := 30.0, [30].Setpoint[53] := 5.0, [30].Setpoint[54] := 5.0, [30].Setpoint[55] := 3.0, [30].Setpoint[57] := 300.0, [30].Name := 'RECIPE #30', [31].Setpoint[1] := 55.0, [31].Setpoint[2] := 65.0, [31].Setpoint[3] := 60.0, [31].Setpoint[4] := 45.0, [31].Setpoint[5] := 65.0, [31].Setpoint[7] := 53.0, [31].Setpoint[8] := 63.0, [31].Setpoint[9] := 57.0, [31].Setpoint[10] := 43.0, [31].Setpoint[11] := 63.0, [31].Setpoint[13] := 85.0, [31].Setpoint[14] := 300.0, [31].Setpoint[15] := 900.0, [31].Setpoint[17] := 15.0, [31].Setpoint[18] := 14.0, [31].Setpoint[19] := 15.0, [31].Setpoint[20] := 45.0, [31].Setpoint[21] := 5.0, [31].Setpoint[22] := 15.0, [31].Setpoint[23] := 300.0, [31].Setpoint[25] := 10.0, [31].Setpoint[26] := 9.0, [31].Setpoint[27] := 10.0, [31].Setpoint[28] := 50.0, [31].Setpoint[29] := 3.0, [31].Setpoint[30] := 17.0, [31].Setpoint[31] := 300.0, [31].Setpoint[33] := 2.0, [31].Setpoint[34] := 900.0, [31].Setpoint[37] := 35.0, [31].Setpoint[41] := 5.0, [31].Setpoint[42] := 50.0,
        [31].Setpoint[43] := 5.0, [31].Setpoint[44] := 60.0, [31].Setpoint[45] := 50.0, [31].Setpoint[47] := 15.0, [31].Setpoint[49] := 180.0, [31].Setpoint[50] := 180.0, [31].Setpoint[52] := 30.0, [31].Setpoint[53] := 5.0, [31].Setpoint[54] := 5.0, [31].Setpoint[55] := 3.0, [31].Setpoint[57] := 300.0, [31].Name := 'RECIPE #31', [32].Setpoint[1] := 55.0, [32].Setpoint[2] := 65.0, [32].Setpoint[3] := 60.0, [32].Setpoint[4] := 45.0, [32].Setpoint[5] := 65.0, [32].Setpoint[7] := 53.0, [32].Setpoint[8] := 63.0, [32].Setpoint[9] := 57.0, [32].Setpoint[10] := 43.0, [32].Setpoint[11] := 63.0, [32].Setpoint[13] := 85.0, [32].Setpoint[14] := 300.0, [32].Setpoint[15] := 900.0, [32].Setpoint[17] := 15.0, [32].Setpoint[18] := 14.0, [32].Setpoint[19] := 15.0, [32].Setpoint[20] := 45.0, [32].Setpoint[21] := 5.0, [32].Setpoint[22] := 15.0, [32].Setpoint[23] := 300.0, [32].Setpoint[25] := 10.0, [32].Setpoint[26] := 9.0, [32].Setpoint[27] := 10.0, [32].Setpoint[28] := 50.0, [32].Setpoint[29] := 3.0, [32].Setpoint[30] := 17.0, [32].Setpoint[31] := 300.0, [32].Setpoint[33] := 2.0, [32].Setpoint[34] := 900.0, [32].Setpoint[37] := 35.0, [32].Setpoint[41] := 5.0, [32].Setpoint[42] := 50.0, [32].Setpoint[43] := 5.0, [32].Setpoint[44] := 60.0, [32].Setpoint[45] := 50.0, [32].Setpoint[47] := 15.0, [32].Setpoint[49] := 180.0, [32].Setpoint[50] := 180.0, [32].Setpoint[52] := 30.0, [32].Setpoint[53] := 5.0, [32].Setpoint[54] := 5.0, [32].Setpoint[55] := 3.0, [32].Setpoint[57] := 300.0, [32].Name := 'RECIPE #32', [33].Setpoint[1] := 55.0, [33].Setpoint[2] := 65.0, [33].Setpoint[3] := 60.0, [33].Setpoint[4] := 45.0,
        [33].Setpoint[5] := 65.0, [33].Setpoint[7] := 53.0, [33].Setpoint[8] := 63.0, [33].Setpoint[9] := 57.0, [33].Setpoint[10] := 43.0, [33].Setpoint[11] := 63.0, [33].Setpoint[13] := 85.0, [33].Setpoint[14] := 300.0, [33].Setpoint[15] := 900.0, [33].Setpoint[17] := 15.0, [33].Setpoint[18] := 14.0, [33].Setpoint[19] := 15.0, [33].Setpoint[20] := 45.0, [33].Setpoint[21] := 5.0, [33].Setpoint[22] := 15.0, [33].Setpoint[23] := 300.0, [33].Setpoint[25] := 10.0, [33].Setpoint[26] := 9.0, [33].Setpoint[27] := 10.0, [33].Setpoint[28] := 50.0, [33].Setpoint[29] := 3.0, [33].Setpoint[30] := 17.0, [33].Setpoint[31] := 300.0, [33].Setpoint[33] := 2.0, [33].Setpoint[34] := 900.0, [33].Setpoint[37] := 35.0, [33].Setpoint[41] := 5.0, [33].Setpoint[42] := 50.0, [33].Setpoint[43] := 5.0, [33].Setpoint[44] := 60.0, [33].Setpoint[45] := 50.0, [33].Setpoint[47] := 15.0, [33].Setpoint[49] := 180.0, [33].Setpoint[50] := 180.0, [33].Setpoint[52] := 30.0, [33].Setpoint[53] := 5.0, [33].Setpoint[54] := 5.0, [33].Setpoint[55] := 3.0, [33].Setpoint[57] := 300.0, [33].Name := 'RECIPE #33', [34].Setpoint[1] := 55.0, [34].Setpoint[2] := 65.0, [34].Setpoint[3] := 60.0, [34].Setpoint[4] := 45.0, [34].Setpoint[5] := 65.0, [34].Setpoint[7] := 53.0, [34].Setpoint[8] := 63.0, [34].Setpoint[9] := 57.0, [34].Setpoint[10] := 43.0, [34].Setpoint[11] := 63.0, [34].Setpoint[13] := 85.0, [34].Setpoint[14] := 300.0, [34].Setpoint[15] := 900.0, [34].Setpoint[17] := 15.0, [34].Setpoint[18] := 14.0, [34].Setpoint[19] := 15.0, [34].Setpoint[20] := 45.0, [34].Setpoint[21] := 5.0, [34].Setpoint[22] := 15.0, [34].Setpoint[23] := 300.0,
        [34].Setpoint[25] := 10.0, [34].Setpoint[26] := 9.0, [34].Setpoint[27] := 10.0, [34].Setpoint[28] := 50.0, [34].Setpoint[29] := 3.0, [34].Setpoint[30] := 17.0, [34].Setpoint[31] := 300.0, [34].Setpoint[33] := 2.0, [34].Setpoint[34] := 900.0, [34].Setpoint[37] := 35.0, [34].Setpoint[41] := 5.0, [34].Setpoint[42] := 50.0, [34].Setpoint[43] := 5.0, [34].Setpoint[44] := 60.0, [34].Setpoint[45] := 50.0, [34].Setpoint[47] := 15.0, [34].Setpoint[49] := 180.0, [34].Setpoint[50] := 180.0, [34].Setpoint[52] := 30.0, [34].Setpoint[53] := 5.0, [34].Setpoint[54] := 5.0, [34].Setpoint[55] := 3.0, [34].Setpoint[57] := 300.0, [34].Name := 'RECIPE #34', [35].Setpoint[1] := 55.0, [35].Setpoint[2] := 65.0, [35].Setpoint[3] := 60.0, [35].Setpoint[4] := 45.0, [35].Setpoint[5] := 65.0, [35].Setpoint[7] := 53.0, [35].Setpoint[8] := 63.0, [35].Setpoint[9] := 57.0, [35].Setpoint[10] := 43.0, [35].Setpoint[11] := 63.0, [35].Setpoint[13] := 85.0, [35].Setpoint[14] := 300.0, [35].Setpoint[15] := 900.0, [35].Setpoint[17] := 15.0, [35].Setpoint[18] := 14.0, [35].Setpoint[19] := 15.0, [35].Setpoint[20] := 45.0, [35].Setpoint[21] := 5.0, [35].Setpoint[22] := 15.0, [35].Setpoint[23] := 300.0, [35].Setpoint[25] := 10.0, [35].Setpoint[26] := 9.0, [35].Setpoint[27] := 10.0, [35].Setpoint[28] := 50.0, [35].Setpoint[29] := 3.0, [35].Setpoint[30] := 17.0, [35].Setpoint[31] := 300.0, [35].Setpoint[33] := 2.0, [35].Setpoint[34] := 900.0, [35].Setpoint[37] := 35.0, [35].Setpoint[41] := 5.0, [35].Setpoint[42] := 50.0, [35].Setpoint[43] := 5.0, [35].Setpoint[44] := 60.0, [35].Setpoint[45] := 50.0, [35].Setpoint[47] := 15.0,
        [35].Setpoint[49] := 180.0, [35].Setpoint[50] := 180.0, [35].Setpoint[52] := 30.0, [35].Setpoint[53] := 5.0, [35].Setpoint[54] := 5.0, [35].Setpoint[55] := 3.0, [35].Setpoint[57] := 300.0, [35].Name := 'RECIPE #35', [36].Setpoint[1] := 55.0, [36].Setpoint[2] := 65.0, [36].Setpoint[3] := 60.0, [36].Setpoint[4] := 45.0, [36].Setpoint[5] := 65.0, [36].Setpoint[7] := 53.0, [36].Setpoint[8] := 63.0, [36].Setpoint[9] := 57.0, [36].Setpoint[10] := 43.0, [36].Setpoint[11] := 63.0, [36].Setpoint[13] := 85.0, [36].Setpoint[14] := 300.0, [36].Setpoint[15] := 900.0, [36].Setpoint[17] := 15.0, [36].Setpoint[18] := 14.0, [36].Setpoint[19] := 15.0, [36].Setpoint[20] := 45.0, [36].Setpoint[21] := 5.0, [36].Setpoint[22] := 15.0, [36].Setpoint[23] := 300.0, [36].Setpoint[25] := 10.0, [36].Setpoint[26] := 9.0, [36].Setpoint[27] := 10.0, [36].Setpoint[28] := 50.0, [36].Setpoint[29] := 3.0, [36].Setpoint[30] := 17.0, [36].Setpoint[31] := 300.0, [36].Setpoint[33] := 2.0, [36].Setpoint[34] := 900.0, [36].Setpoint[37] := 35.0, [36].Setpoint[41] := 5.0, [36].Setpoint[42] := 50.0, [36].Setpoint[43] := 5.0, [36].Setpoint[44] := 60.0, [36].Setpoint[45] := 50.0, [36].Setpoint[47] := 15.0, [36].Setpoint[49] := 180.0, [36].Setpoint[50] := 180.0, [36].Setpoint[52] := 30.0, [36].Setpoint[53] := 5.0, [36].Setpoint[54] := 5.0, [36].Setpoint[55] := 3.0, [36].Setpoint[57] := 300.0, [36].Name := 'RECIPE #36', [37].Setpoint[1] := 55.0, [37].Setpoint[2] := 65.0, [37].Setpoint[3] := 60.0, [37].Setpoint[4] := 45.0, [37].Setpoint[5] := 65.0, [37].Setpoint[7] := 53.0, [37].Setpoint[8] := 63.0, [37].Setpoint[9] := 57.0,
        [37].Setpoint[10] := 43.0, [37].Setpoint[11] := 63.0, [37].Setpoint[13] := 85.0, [37].Setpoint[14] := 300.0, [37].Setpoint[15] := 900.0, [37].Setpoint[17] := 15.0, [37].Setpoint[18] := 14.0, [37].Setpoint[19] := 15.0, [37].Setpoint[20] := 45.0, [37].Setpoint[21] := 5.0, [37].Setpoint[22] := 15.0, [37].Setpoint[23] := 300.0, [37].Setpoint[25] := 10.0, [37].Setpoint[26] := 9.0, [37].Setpoint[27] := 10.0, [37].Setpoint[28] := 50.0, [37].Setpoint[29] := 3.0, [37].Setpoint[30] := 17.0, [37].Setpoint[31] := 300.0, [37].Setpoint[33] := 2.0, [37].Setpoint[34] := 900.0, [37].Setpoint[37] := 35.0, [37].Setpoint[41] := 5.0, [37].Setpoint[42] := 50.0, [37].Setpoint[43] := 5.0, [37].Setpoint[44] := 60.0, [37].Setpoint[45] := 50.0, [37].Setpoint[47] := 15.0, [37].Setpoint[49] := 180.0, [37].Setpoint[50] := 180.0, [37].Setpoint[52] := 30.0, [37].Setpoint[53] := 5.0, [37].Setpoint[54] := 5.0, [37].Setpoint[55] := 3.0, [37].Setpoint[57] := 300.0, [37].Name := 'RECIPE #37', [38].OpCode[1] := 4, [38].OpCode[2] := 8, [38].OpCode[3] := 7, [38].OpCode[4] := 13, [38].OpCode[5] := 5, [38].OpCode[6] := 2, [38].OpCode[7] := 1, [38].StepTime[1] := 10, [38].StepTime[2] := 20, [38].StepTime[3] := 10, [38].StepTime[4] := 20, [38].StepTime[5] := 10, [38].StepTime[6] := 10, [38].StepTime[7] := 10, [38].Setpoint[1] := 20.0, [38].Setpoint[2] := 90.0, [38].Setpoint[3] := 60.0, [38].Setpoint[4] := 45.0, [38].Setpoint[5] := 65.0, [38].Setpoint[7] := 20.0, [38].Setpoint[8] := 85.0, [38].Setpoint[9] := 57.0, [38].Setpoint[10] := 43.0, [38].Setpoint[11] := 63.0,
        [38].Setpoint[13] := 95.0, [38].Setpoint[14] := 9999.0, [38].Setpoint[15] := 9999.0, [38].Setpoint[17] := 15.0, [38].Setpoint[18] := 14.0, [38].Setpoint[19] := 15.0, [38].Setpoint[20] := 45.0, [38].Setpoint[21] := 5.0, [38].Setpoint[22] := 15.0, [38].Setpoint[23] := 300.0, [38].Setpoint[25] := 10.0, [38].Setpoint[26] := 9.0, [38].Setpoint[27] := 10.0, [38].Setpoint[28] := 50.0, [38].Setpoint[29] := 3.0, [38].Setpoint[30] := 17.0, [38].Setpoint[31] := 300.0, [38].Setpoint[33] := 2.0, [38].Setpoint[34] := 900.0, [38].Setpoint[37] := 45.0, [38].Setpoint[41] := 5.0, [38].Setpoint[42] := 60.0, [38].Setpoint[43] := 5.0, [38].Setpoint[44] := 100.0, [38].Setpoint[45] := 50.0, [38].Setpoint[47] := 15.0, [38].Setpoint[49] := 180.0, [38].Setpoint[50] := 180.0, [38].Setpoint[52] := 30.0, [38].Setpoint[53] := 5.0, [38].Setpoint[54] := 5.0, [38].Setpoint[55] := 3.0, [38].Setpoint[57] := 300.0, [38].Name := 'SYSTEM PERFORMANCE', [39].OpCode[1] := 4, [39].OpCode[2] := 8, [39].OpCode[3] := 9, [39].OpCode[4] := 5, [39].OpCode[5] := 4, [39].OpCode[6] := 7, [39].OpCode[7] := 10, [39].OpCode[8] := 13, [39].OpCode[9] := 16, [39].OpCode[10] := 20, [39].OpCode[11] := 5, [39].OpCode[12] := 4, [39].OpCode[13] := 11, [39].OpCode[14] := 13, [39].OpCode[15] := 16, [39].OpCode[16] := 14, [39].OpCode[17] := 17, [39].OpCode[18] := 18, [39].OpCode[19] := 2, [39].OpCode[20] := 1, [39].StepTime[1] := 10, [39].StepTime[2] := 10, [39].StepTime[3] := 10, [39].StepTime[4] := 10, [39].StepTime[5] := 10, [39].StepTime[6] := 10,
        [39].StepTime[7] := 10, [39].StepTime[8] := 10, [39].StepTime[9] := 10, [39].StepTime[10] := 10, [39].StepTime[11] := 10, [39].StepTime[12] := 10, [39].StepTime[13] := 10, [39].StepTime[14] := 10, [39].StepTime[15] := 10, [39].StepTime[16] := 10, [39].StepTime[17] := 10, [39].StepTime[18] := 10, [39].StepTime[19] := 10, [39].StepTime[20] := 10, [39].Setpoint[1] := 55.0, [39].Setpoint[2] := 65.0, [39].Setpoint[3] := 60.0, [39].Setpoint[4] := 45.0, [39].Setpoint[5] := 65.0, [39].Setpoint[7] := 53.0, [39].Setpoint[8] := 63.0, [39].Setpoint[9] := 57.0, [39].Setpoint[10] := 43.0, [39].Setpoint[11] := 63.0, [39].Setpoint[13] := 85.0, [39].Setpoint[14] := 300.0, [39].Setpoint[15] := 900.0, [39].Setpoint[17] := 15.0, [39].Setpoint[18] := 14.0, [39].Setpoint[19] := 15.0, [39].Setpoint[20] := 45.0, [39].Setpoint[21] := 5.0, [39].Setpoint[22] := 15.0, [39].Setpoint[23] := 300.0, [39].Setpoint[25] := 10.0, [39].Setpoint[26] := 9.0, [39].Setpoint[27] := 10.0, [39].Setpoint[28] := 50.0, [39].Setpoint[29] := 3.0, [39].Setpoint[30] := 17.0, [39].Setpoint[31] := 300.0, [39].Setpoint[33] := 2.0, [39].Setpoint[34] := 900.0, [39].Setpoint[37] := 35.0, [39].Setpoint[41] := 5.0, [39].Setpoint[42] := 50.0, [39].Setpoint[43] := 5.0, [39].Setpoint[44] := 60.0, [39].Setpoint[45] := 50.0, [39].Setpoint[47] := 15.0, [39].Setpoint[49] := 180.0, [39].Setpoint[50] := 180.0, [39].Setpoint[52] := 30.0, [39].Setpoint[53] := 5.0, [39].Setpoint[54] := 5.0, [39].Setpoint[55] := 3.0, [39].Setpoint[57] := 300.0, [39].Name := 'FAT TEST RECIPE', [40].OpCode[1] := 2, [40].OpCode[2] := 4,
        [40].OpCode[3] := 13, [40].OpCode[4] := 5, [40].OpCode[5] := 2, [40].OpCode[6] := 1, [40].StepTime[1] := 10, [40].StepTime[2] := 10, [40].StepTime[3] := 10, [40].StepTime[4] := 10, [40].StepTime[5] := 10, [40].StepTime[6] := 10, [40].Setpoint[1] := 55.0, [40].Setpoint[2] := 65.0, [40].Setpoint[3] := 60.0, [40].Setpoint[4] := 45.0, [40].Setpoint[5] := 65.0, [40].Setpoint[7] := 53.0, [40].Setpoint[8] := 63.0, [40].Setpoint[9] := 57.0, [40].Setpoint[10] := 43.0, [40].Setpoint[11] := 63.0, [40].Setpoint[13] := 85.0, [40].Setpoint[14] := 300.0, [40].Setpoint[15] := 900.0, [40].Setpoint[17] := 15.0, [40].Setpoint[18] := 14.0, [40].Setpoint[19] := 15.0, [40].Setpoint[20] := 45.0, [40].Setpoint[21] := 5.0, [40].Setpoint[22] := 15.0, [40].Setpoint[23] := 300.0, [40].Setpoint[25] := 10.0, [40].Setpoint[26] := 9.0, [40].Setpoint[27] := 10.0, [40].Setpoint[28] := 50.0, [40].Setpoint[29] := 3.0, [40].Setpoint[30] := 17.0, [40].Setpoint[31] := 300.0, [40].Setpoint[33] := 2.0, [40].Setpoint[34] := 900.0, [40].Setpoint[37] := 35.0, [40].Setpoint[41] := 5.0, [40].Setpoint[42] := 50.0, [40].Setpoint[43] := 5.0, [40].Setpoint[44] := 60.0, [40].Setpoint[45] := 50.0, [40].Setpoint[47] := 15.0, [40].Setpoint[49] := 180.0, [40].Setpoint[50] := 180.0, [40].Setpoint[52] := 30.0, [40].Setpoint[53] := 5.0, [40].Setpoint[54] := 5.0, [40].Setpoint[55] := 3.0, [40].Setpoint[57] := 300.0, [40].Name := 'SEPARATOR TANK FLUSH');   // RECIPES
        [0].Setpoint[0]   // CURRENT RECIPE SETPOINTS
        [0].Setpoint[16]   // MASTER SETPOINT
        [0].Setpoint[24]   // MASTER SETPOINT
        [0].Setpoint[32]   // MASTER SETPOINT
        [0].Setpoint[35]   // MASTER SETPOINT
        [0].Setpoint[36]   // MASTER SETPOINT
        [0].Setpoint[13]   // MASTER SETPOINT HIGH SUPPLY TEMPERATURE
        [0].Setpoint[10]   // MASTER SETPOINT RETURN TEMP 4 (CHEM #2 WASH)
        [0].Setpoint[38]   // MASTER SETPOINT
        [0].Setpoint[49]   // MASTER SETPOINT SEPARATOR FILL HOLD WATCHDOG
        [0].Setpoint[6]   // MASTER SETPOINT
        [0].Setpoint[12]   // MASTER SETPOINT
        [0].Setpoint[46]   // MASTER SETPOINT
        [0].Setpoint[20]   // MASTER SETPOINT CHEM #1 MIX TIME
        [0].Setpoint[61]   // MASTER SETPOINT
        [0].Setpoint[33]   // MASTER SETPOINT RINSE CONDUCTIVITY
        [0].Setpoint[48]   // MASTER SETPOINT
        [0].Setpoint[51]   // MASTER SETPOINT
        [0].Setpoint[59]   // MASTER SETPOINT
        [0].Setpoint[3]   // MASTER SETPOINT SUPPLY TEMP 3 (CHEM #1 WASH)
        [0].Setpoint[11]   // MASTER SETPOINT RETURN TEMP 5 (FINAL RINSE)
        [0].Setpoint[44]   // MASTER SETPOINT HIGH SUPPLY PRESSURE ALARM
        [0].Setpoint[1]   // MASTER SETPOINT SUPPLY TEMP 1 (PRE-RINSE)
        [0].Setpoint[39]   // MASTER SETPOINT
        [0].Setpoint[45]   // MASTER SETPOINT PUMP TO DRAIN FLOW MODULATION
        [0].Setpoint[40]   // MASTER SETPOINT
        [0].Setpoint[60]   // MASTER SETPOINT
        [0].Setpoint[62]   // MASTER SETPOINT
        [0].Setpoint[28]   // MASTER SETPOINT CHEM #2 MIX TIME
        [0].Setpoint[63]   // MASTER SETPOINT
        [0].Setpoint[64]   // MASTER SETPOINT
        [0].Setpoint[7]   // MASTER SETPOINT RETURN TEMP 1 (PRE-RINSE)
        [0].Setpoint[19]   // MASTER SETPOINT CHEM #1 PUMP INJECTION TIME
        [0].Setpoint[50]   // MASTER SETPOINT SEPARATOR EMPTY HOLD WATCHDOG
        [0].Setpoint[27]   // MASTER SETPOINT CHEM #2 PUMP INJECTION TIME
        [0].Setpoint[58]   // MASTER SETPOINT
        [0].Setpoint[53]   // MASTER SETPOINT SUPPLY FLOW VALVE POSITION DEADBAND
        [0].Setpoint[65]   // MASTER SETPOINT
        [0].Setpoint[2]   // MASTER SETPOINT SUPPLY TEMP 2 (RINSE)
        [0].Setpoint[66]   // MASTER SETPOINT
        [0].Setpoint[67]   // MASTER SETPOINT
        [0].Setpoint[37]   // MASTER SETPOINT SUPPLY FLOW RATE
        [0].Setpoint[8]   // MASTER SETPOINT RETURN TEMP 2 (RINSE)
        [0].Setpoint[75]   // MASTER SETPOINT
        [0].Setpoint[76]   // MASTER SETPOINT
        [0].Setpoint[14]   // MASTER SETPOINT SUPPLY TEMPERATURE HOLD WATCHDOG
        [0].Setpoint[22]   // MASTER SETPOINT CHEM #1 PUMP BURST OFF
        [0].Setpoint[57]   // MASTER SETPOINT OVERFLOW TANK EMPTY HOLD WATCHDOG
        [0].Setpoint[68]   // MASTER SETPOINT
        [0].Setpoint[69]   // MASTER SETPOINT
        [0].Setpoint[70]   // MASTER SETPOINT
        [0].Setpoint[71]   // MASTER SETPOINT
        [0].Setpoint[72]   // MASTER SETPOINT
        [0].Setpoint[73]   // MASTER SETPOINT
        [0].Setpoint[21]   // MASTER SETPOINT CHEM #1 PUMP BURST ON
        [0].Setpoint[74]   // MASTER SETPOINT
        [0].Setpoint[23]   // MASTER SETPOINT CHEM #1 CONDUCTIVITY HOLD WATCHDOG
        [0].Setpoint[18]   // MASTER SETPOINT CHEM #1 CONDUCTIVITY HOLD
        [0].Setpoint[77]   // MASTER SETPOINT
        [0].Setpoint[78]   // MASTER SETPOINT
        [0].Setpoint[29]   // MASTER SETPOINT CHEM #2 PUMP BURST ON
        [0].Setpoint[79]   // MASTER SETPOINT
        [0].Setpoint[47]   // MASTER SETPOINT AWFI DRAIN FLOW MODULATION
        [0].Setpoint[15]   // MASTER SETPOINT RETURN TEMPERATURE HOLD WATCHDOG
        [0].Setpoint[31]   // MASTER SETPOINT CHEM #2 CONDUCTIVITY HOLD WATCHDOG
        [0].Setpoint[81]   // MASTER SETPOINT
        [0].Setpoint[30]   // MASTER SETPOINT CHEM #2 PUMP BURST OFF
        [0].Setpoint[41]   // MASTER SETPOINT LOW SUPPLY FLOW ALARM
        [0].Setpoint[17]   // MASTER SETPOINT CHEM #1 CONDUCTIVITY
        [0].Setpoint[9]   // MASTER SETPOINT RETURN TEMP 3 (CHEM #1 WASH)
        [0].Setpoint[4]   // MASTER SETPOINT SUPPLY TEMP 4 (CHEM #2 WASH)
        [0].Setpoint[80]   // MASTER SETPOINT
        [0].Setpoint[82]   // MASTER SETPOINT
        [0].Setpoint[83]   // MASTER SETPOINT
        [0].Setpoint[26]   // MASTER SETPOINT CHEM #2 CONDUCTIVITY HOLD
        [0].Setpoint[84]   // MASTER SETPOINT
        [0].Setpoint[42]   // MASTER SETPOINT HIGH SUPPLY FLOW ALARM
        [0].Setpoint[34]   // MASTER SETPOINT RINSE CONDUCTIVITY HOLD WATCHDOG
        [0].Setpoint[52]   // MASTER SETPOINT SEPARATOR LOW LEVEL SHUTDOWN DELAY
        [0].Setpoint[55]   // MASTER SETPOINT OVERFLOW TANK DRAIN PUMP DELAY
        [0].Setpoint[54]   // MASTER SETPOINT DRAIN FLOW VALVE POSITION DEADBAND
        [0].Setpoint[43]   // MASTER SETPOINT LOW SUPPLY PRESSURE ALARM
        [0].Setpoint[56]   // MASTER SETPOINT PROCESS EQUIPMENT INTERFACE ENABLE
        [0].Setpoint[85]   // MASTER SETPOINT
        [0].Setpoint[5]   // MASTER SETPOINT SUPPLY TEMP 5 (FINAL RINSE)
        [0].Setpoint[25]   // MASTER SETPOINT CHEM #2 CONDUCTIVITY
        [0].Setpoint[86]   // MASTER SETPOINT
        [0].Setpoint[87]   // MASTER SETPOINT
        [0].Setpoint[88]   // MASTER SETPOINT
        [0].Setpoint[89]   // MASTER SETPOINT
        [0].Setpoint[90]   // MASTER SETPOINT
        [0].Setpoint[91]   // MASTER SETPOINT
        [0].Setpoint[92]   // MASTER SETPOINT
        [0].Setpoint[93]   // MASTER SETPOINT
        [0].Setpoint[94]   // MASTER SETPOINT
        [0].Setpoint[95]   // MASTER SETPOINT
        [0].Setpoint[96]   // MASTER SETPOINT
   Recipe_Name : STRING[41] := ([1] := 'WASH CYCLE', [2] := 'RECIPE #2', [3] := 'RECIPE #3', [4] := 'RECIPE #4', [5] := 'RECIPE #5', [6] := 'RECIPE #6', [7] := 'RECIPE #7', [8] := 'RECIPE #8', [9] := 'RECIPE #9', [10] := 'RECIPE #10', [11] := 'RECIPE #11', [12] := 'RECIPE #12', [13] := 'RECIPE #13', [14] := 'RECIPE #14', [15] := 'RECIPE #15', [16] := 'RECIPE #16', [17] := 'RECIPE #17', [18] := 'RECIPE #18', [19] := 'RECIPE #19', [20] := 'RECIPE #20', [21] := 'RECIPE #21', [22] := 'RECIPE #22', [23] := 'RECIPE #23', [24] := 'RECIPE #24', [25] := 'RECIPE #25', [26] := 'RECIPE #26', [27] := 'RECIPE #27', [28] := 'RECIPE #28', [29] := 'RECIPE #29', [30] := 'RECIPE #30', [31] := 'RECIPE #31', [32] := 'RECIPE #32', [33] := 'RECIPE #33', [34] := 'RECIPE #34', [35] := 'RECIPE #35', [36] := 'RECIPE #36', [37] := 'RECIPE #37', [38] := 'SYSTEM PERFORMANCE', [39] := 'FAT TEST RECIPE', [40] := 'SEPARATOR TANK FLUSH');   // RECIPE NAME STORAGE
   Recipe_Name_Indx : DINT := 3;   // RECIPE NAME INDEX POSITION
   Recipe_Step_Length : CONTROL := (LEN := 97, POS := 20, EN := 1, IN := 1, FD := 1);   // CURRENT RECIPE LENGTH
   SCLD_Drain_Flow : SCALE := (InRawMax := 100.0, InEUMax := 16383.0);   // DRAIN FLOW MODULATION 0-100%
   SCLD_DrainValve_Feedback : SCALE := (In := 3132.0, InRawMax := 16383.0, InRawMin := 3277.0, InEUMax := 100.0, Out := -1.1063635, MinAlarm := 1);   // DRAIN FLOW FEEDBACK POSITION 0-100%
   SCLD_Return_Temp : SCALE := (In := 6183.0, InRawMax := 16383.0, InRawMin := 3277.0, InEUMax := 100.0, Out := 22.17305);   // RETURN TEMPERATURE 0-100°C
   SCLD_Rinse_Cond : SCALE := (In := 4799.0, InRawMax := 16383.0, InRawMin := 3277.0, InEUMax := 10.0, Limiting := 1, Out := 1.1613002);   // RINSE CONDUCTIVITY 0-10 uS/cm
   SCLD_Spare_IN_264 : SCALE := (In := -8.0, InRawMax := 16383.0, InRawMin := 3277.0, InEUMax := 100.0, Out := -25.064856, MinAlarm := 1);   // SPARE IN-264
   SCLD_Spare_IN_272 : SCALE := (In := -9.0, InRawMax := 16383.0, InRawMin := 3277.0, InEUMax := 100.0, Out := -25.072485, MinAlarm := 1);   // SPARE IN-272
   SCLD_Supply_Flow : SCALE := (In := 3267.0, InRawMax := 16383.0, InRawMin := 3277.0, InEUMax := 60.0, Limiting := 1, MinAlarm := 1);   // SUPPLY FLOW 0-60 GPM
   SCLD_Supply_Press : SCALE := (In := 3256.0, InRawMax := 16383.0, InRawMin := 3277.0, InEUMax := 100.0, Limiting := 1, MinAlarm := 1);   // SUPPLY PRESSURE 0-100 PSIG
   SCLD_Supply_Temp : SCALE := (In := 6166.0, InRawMax := 16383.0, InRawMin := 3277.0, InEUMax := 100.0, Out := 22.043339);   // SUPPLY TEMPERATURE 0-100°C
   SCLD_SupplyValve_Feedback : SCALE := (In := 3173.0, InRawMax := 16383.0, InRawMin := 3277.0, InEUMax := 100.0, Out := -0.7935297, MinAlarm := 1);   // SUPPLY FLOW FEEDBACK POSITION 0-100%
   SCLD_Wash_Cond : SCALE := (In := 3260.0, InRawMax := 16383.0, InRawMin := 3277.0, InEUMax := 100.0, Limiting := 1, MinAlarm := 1);   // WASH CONDUCTIVITY 0-100 mS/cm
   SecurityLevel : DINT := 2;   // MAIN HMI CURRENT LOGGED IN OPERATOR
   Sequencer : CONTROL[4] := ([0].LEN := 97, [1].LEN := 97, [1].EN := 1, [2].LEN := 97, [2].POS := 9, [2].EN := 1, [3].LEN := 1, [3].POS := 1, [3].DN := 1);   // SEQUENCER
        [0]   // MASTER RECIPE STEP SEQUENCER
        [3]   // MESSAGE SEQUENCER
        [2]   // SUBSEQUENT STEP OPCODE SEQUENCER
        [1]   // CURRENT OPCODE SEQUENCER
   SP_Drain_Flow : REAL;   // CURRENT DRAIN FLOW MODULATION SETPOINT
   SP_DrainValve_HighDeadband : REAL := 5.0;   // CURRENT DRAIN VALVE DEADBAND SETPOINT
   SP_DrainValve_LowDeadband : REAL := -5.0;   // CURRENT DRAIN VALVE DEADBAND SETPOINT
   SP_Return_Temp : REAL;   // CURRENT RETURN TEMP SETPOINT
   SP_Rinse_Cond : REAL;   // CURRENT RINSE CONDUCTIVITY SETPOINT
   SP_Supply_Flow : REAL;   // CURRENT SUPPLY FLOW SETPOINT
   SP_Supply_Temp : REAL;   // CURRENT SUPPLY TEMP SETPOINT
   SP_SupplyValve_HighDeadband : REAL := 5.0;   // CURRENT SUPPLY VALVE DEADBAND SETPOINT
   SP_SupplyValve_LowDeadband : REAL := -5.0;   // CURRENT SUPPLY VALVE DEADBAND SETPOINT
   SP_Wash_Cond : REAL;   // CURRENT WASH CONDUCTIVITY SETPOINT
   SP_Wash_Cond_Hold : REAL;   // CURRENT WASH CONDUCTIVITY SETPOINT LOW HOLD
   Step_Time_Min : STRING := '0';
   Step_Time_Preset : DINT;
   Step_Time_Remaining : STRING[5] := ([0] := '0:0', [1] := '0:00', [2] := ':', [3] := ':0');
   Step_Time_Sec : STRING := '0';
   Subsequent_OpCode_Pin : DINT[5] := ([1] := 21, [2] := 43008);   // OPCODE PIN ARRAY
        [2]   // SEQUENCER OUTPUTS WORD #2
        [3]   // SEQUENCER OUTPUTS WORD #3
        [4]   // SEQUENCER OUTPUTS WORD #4
        [3].0   // SEQ PIN WORD #3 PIN #00
        [3].1   // SEQ PIN WORD #3 PIN #01
        [3].2   // SEQ PIN WORD #3 PIN #02
        [1].2   // SEQ PIN WORD #1 PIN #02
        [1].8   // SEQ PIN WORD #1 PIN #08
        [2].2   // SEQ PIN WORD #2 PIN #02
        [3].3   // SEQ PIN WORD #3 PIN #03
        [3].4   // SEQ PIN WORD #3 PIN #04
        [3].5   // SEQ PIN WORD #3 PIN #05
        [3].9   // SEQ PIN WORD #3 PIN #09
        [1]   // SEQUENCER OUTPUTS WORD #1
        [1].0   // SEQ PIN WORD #1 PIN #00 WFI FILL ON
        [1].1   // SEQ PIN WORD #1 PIN #01 PW FILL ON
        [2].3   // SEQ PIN WORD #2 PIN #03
        [1].13   // SEQ PIN WORD #1 PIN #13 FILL HOLD
        [1].14   // SEQ PIN WORD #1 PIN #14
        [1].3   // SEQ PIN WORD #1 PIN #03 PAUSE
        [1].7   // SEQ PIN WORD #1 PIN #07 AIR BLOW
        [1].9   // SEQ PIN WORD #1 PIN #09 EMPTY HOLD
        [2].12   // SEQ PIN WORD #2 PIN #12
        [2].14   // SEQ PIN WORD #2 PIN #14
        [2].4   // SEQ PIN WORD #2 PIN #04 PRE-HEAT
        [2].5   // SEQ PIN WORD #2 PIN #05
        [3].10   // SEQ PIN WORD #3 PIN #10
        [3].11   // SEQ PIN WORD #3 PIN #11
        [3].12   // SEQ PIN WORD #3 PIN #12
        [3].13   // SEQ PIN WORD #3 PIN #13
        [3].14   // SEQ PIN WORD #3 PIN #14
        [3].15   // SEQ PIN WORD #3 PIN #15
        [4].0   // SEQ PIN WORD #4 PIN #00
        [4].1   // SEQ PIN WORD #4 PIN #01
        [4].10   // SEQ PIN WORD #4 PIN #10
        [4].11   // SEQ PIN WORD #4 PIN #11
        [4].12   // SEQ PIN WORD #4 PIN #12
        [4].13   // SEQ PIN WORD #4 PIN #13
        [4].14   // SEQ PIN WORD #4 PIN #14
        [4].15   // SEQ PIN WORD #4 PIN #15
        [4].2   // SEQ PIN WORD #4 PIN #02
        [4].3   // SEQ PIN WORD #4 PIN #03
        [4].4   // SEQ PIN WORD #4 PIN #04
        [4].5   // SEQ PIN WORD #4 PIN #05
        [4].6   // SEQ PIN WORD #4 PIN #06
        [4].7   // SEQ PIN WORD #4 PIN #07
        [1].10   // SEQ PIN WORD #1 PIN #10 RINSE CONDUCTIVITY HOLD
        [1].11   // SEQ PIN WORD #1 PIN #11 WASH CONDUCTIVITY HOLD
        [1].12   // SEQ PIN WORD #1 PIN #12 TEMPERATURE HOLD
        [1].15   // SEQ PIN WORD #1 PIN #15 LOW LEVEL DISABLE
        [1].4   // SEQ PIN WORD #1 PIN #04 MODULATION DRAIN VALVE
        [1].5   // SEQ PIN WORD #1 PIN #05 PUMP CASING DRAIN
        [1].6   // SEQ PIN WORD #1 PIN #06 RETURN LINE DRAIN
        [2].0   // SEQ PIN WORD #2 PIN #00 CHEM #2 CONDUCTIVITY
        [2].1   // SEQ PIN WORD #2 PIN #01 CHEM #1 CONDUCTIVITY
        [2].10   // SEQ PIN WORD #2 PIN #10 TEMP 2 ( RINSE)
        [2].11   // SEQ PIN WORD #2 PIN #11 TEMP 1 (PRE-RINSE)
        [2].13   // SEQ PIN WORD #2 PIN #13 FLOW CONTROL ENABLE
        [2].15   // SEQ PIN WORD #2 PIN #15 SUPPLY PUMP
        [2].6   // SEQ PIN WORD #2 PIN #06 TEMP 6 (SPARE)
        [2].7   // SEQ PIN WORD #2 PIN #07 TEMP 5 (FINAL RINSE)
        [2].8   // SEQ PIN WORD #2 PIN #08 TEMP 4 (CHEM #2 WASH)
        [2].9   // SEQ PIN WORD #2 PIN #09 TEMP 3 (CHEM #1 WASH)
        [3].6   // SEQ PIN WORD #3 PIN #06 PRINT FINAL RINSE CYCLE
        [3].7   // SEQ PIN WORD #3 PIN #07 PRINT CHEM #2 CYCLE
        [3].8   // SEQ PIN WORD #3 PIN #08 PRINT CHEM #1 CYCLE
        [4].8   // SEQ PIN WORD #4 PIN #08
        [4].9   // SEQ PIN WORD #4 PIN #09
   Supply_Mod_Valve_force_open : BOOL;   // FORCE SUPPLY MOD. VALVE TO 100% OPEN
   SYS_Bit : BOOL[128] := ([4] := 1, [6] := 1, [15] := 1, [21] := 1, [25] := 1, [27] := 1, [28] := 1, [30] := 1, [34] := 1, [39] := 1, [40] := 1, [41] := 1, [43] := 1, [64] := 1, [66] := 1, [68] := 1, [81] := 1, [82] := 1, [85] := 1, [87] := 1, [88] := 1);   // SYSTEM BIT
        [46]   // SYSTEM ONE SHOT
   SYS_Timer : TIMER[60] := ([0].PRE := 2000, [0].ACC := 189, [0].EN := 1, [0].TT := 1, [1].PRE := 6000, [2].PRE := 45000, [3].PRE := 75000, [3].ACC := 75000, [3].EN := 1, [3].DN := 1, [4].PRE := 5000, [4].ACC := 5002, [4].EN := 1, [4].DN := 1, [5].PRE := 2000, [6].PRE := 3000, [9].PRE := 3600000, [10].PRE := 3000, [10].ACC := 3000, [10].EN := 1, [10].DN := 1, [11].PRE := 3000, [12].PRE := 3000, [13].PRE := 5000, [14].PRE := 3000, [15].PRE := 3000, [15].ACC := 3000, [15].EN := 1, [15].DN := 1, [16].PRE := 3000, [16].ACC := 3000, [16].EN := 1, [16].DN := 1, [17].PRE := 1, [18].PRE := 3000, [18].ACC := 3000, [18].EN := 1, [18].DN := 1, [20].PRE := 1000, [21].PRE := 3000, [22].PRE := 10000, [22].ACC := 183, [22].EN := 1, [22].TT := 1, [23].PRE := 10000, [24].PRE := 3, [25].PRE := 1000, [26].PRE := 500, [26].ACC := 500, [26].EN := 1, [26].DN := 1, [27].PRE := 20000, [28].PRE := 40000, [29].PRE := 3, [29].ACC := 3, [29].EN := 1, [29].DN := 1, [30].PRE := 1000, [30].ACC := 1001, [30].EN := 1,
        [30].DN := 1, [31].PRE := 1, [32].PRE := 1, [33].PRE := 1, [34].PRE := 1, [35].PRE := 3000, [36].PRE := 20000, [37].PRE := 20000, [38].PRE := 20000, [39].PRE := 20000, [40].PRE := 20, [41].PRE := 20000, [42].PRE := 3000, [42].ACC := 3001, [42].EN := 1, [42].DN := 1, [43].PRE := 3000, [43].ACC := 3001, [43].EN := 1, [43].DN := 1, [44].PRE := 10, [45].PRE := 2, [46].PRE := 10, [46].ACC := 9, [47].PRE := 60000, [48].PRE := 45, [49].PRE := 45000, [50].PRE := 5, [51].PRE := 5, [52].PRE := 3, [52].ACC := 3, [53].PRE := 3, [53].ACC := 1, [55].ACC := 6, [55].EN := 1, [55].DN := 1, [56].PRE := 75, [56].ACC := 75, [57].PRE := 75000, [57].ACC := 75000, [57].EN := 1, [57].DN := 1, [58].PRE := 2000, [59].PRE := 120000);   // SYSTEM TIMER
        [35]   // SYSTEM ALARM ACK ALL DELAY RESET
   TemporaryRecipeSelection : DINT := 39;
   Time_Date : DINT[20] := ([0] := 1998, [1] := 2, [2] := 27, [3] := 5, [4] := 35, [5] := 27, [6] := 287305, [10] := 1998, [11] := 2, [12] := 27, [13] := 5, [14] := 35, [15] := 27, [16] := 287305);   // SYSTEM TIME/DATE EDIT/STORAGE
        [3]   // SYSTEM STORAGE HOUR
        [0]   // SYSTEM STORAGE YEAR
        [2]   // SYSTEM STORAGE DAY
        [13]   // PANELVIEW EDIT HOUR
        [15]   // PANELVIEW EDIT SECONDS
        [5]   // SYSTEM STORAGE SECONDS
        [1]   // SYSTEM STORAGE MONTH
        [11]   // PANELVIEW EDIT MONTH
        [12]   // PANELVIEW EDIT DAY
        [10]   // PANELVIEW EDIT YEAR
        [14]   // PANELVIEW EDIT MINUTE
        [4]   // SYSTEM STORAGE MINUTE
        [6]   // SYSTEM STORAGE MILLISECONDS
   Timer : TIMER[99] := ([0].PRE := 2000, [0].ACC := 1234, [0].EN := 1, [0].TT := 1, [2].PRE := 30000, [3].PRE := 2000, [4].PRE := 1000, [5].PRE := 15000, [6].PRE := 15000, [7].PRE := 3000, [8].PRE := 6000, [9].PRE := 6000, [9].ACC := 6019, [10].PRE := 3000, [10].ACC := 6019, [11].PRE := 6000, [11].ACC := 6000, [11].EN := 1, [11].DN := 1, [12].PRE := 6000, [12].ACC := 6000, [12].EN := 1, [12].DN := 1, [13].PRE := 1000, [14].PRE := 3000, [15].PRE := 3000, [16].PRE := 3000, [16].ACC := 3000, [16].EN := 1, [16].DN := 1, [17].PRE := 1000, [18].PRE := 3000, [18].ACC := 3000, [18].EN := 1, [18].DN := 1, [19].PRE := 5000, [20].PRE := 1000, [20].ACC := 1000, [20].EN := 1, [20].DN := 1, [21].PRE := 3000, [21].ACC := 3000, [22].PRE := 3000, [22].ACC := 3000, [23].PRE := 3, [24].PRE := 3, [25].PRE := 1000, [26].PRE := 20000, [27].PRE := 20000, [28].PRE := 20000, [29].PRE := 3, [29].ACC := 3, [30].PRE := 1000, [31].PRE := 1000, [32].PRE := 1000, [33].PRE := 3000, [34].PRE := 1, [35].PRE := 20000, [36].PRE := 3600000, [36].ACC := 586460,
        [36].EN := 1, [36].TT := 1, [37].PRE := 1500, [38].PRE := 20000, [39].PRE := 45000, [40].PRE := 20, [41].PRE := 2000, [41].ACC := 2000, [42].PRE := 2000, [42].ACC := 2000, [43].PRE := 3000, [43].ACC := 3000, [43].EN := 1, [43].DN := 1, [44].PRE := 10, [45].PRE := 30000, [46].PRE := 15000, [47].PRE := 30000, [48].PRE := 15000, [49].PRE := 45000, [50].PRE := 5, [51].PRE := 5, [52].PRE := 3, [52].ACC := 3, [53].PRE := 3, [53].ACC := 1, [55].PRE := 75000, [55].ACC := 75001, [55].EN := 1, [55].DN := 1, [56].PRE := 75, [56].ACC := 75, [57].PRE := 300000, [58].PRE := 2000, [59].PRE := 120000, [60].PRE := 100, [60].ACC := 58, [63].PRE := 3000, [63].ACC := 3001, [63].EN := 1, [63].DN := 1, [64].PRE := 2000, [64].ACC := 2001, [64].EN := 1, [64].DN := 1, [65].PRE := 2000, [66].PRE := 300000, [68].PRE := 10000, [68].ACC := 964, [68].EN := 1, [68].TT := 1, [70].PRE := 10000, [70].ACC := 966, [70].EN := 1, [70].TT := 1, [74].PRE := 1000, [74].ACC := 1000, [74].EN := 1, [74].DN := 1, [75].PRE := 1000,
        [90].PRE := 5000, [91].PRE := 5000);   // TIMER
        [91]   // RECIPE COMPLETED
        [90]   // RECIPE ABORTED
        [13]   // RINSE CONDUCTIVITY AT SETPOINT DELAY
        [9]   // MANUAL STEP ENABLE DURATION
        [1]   // STEP TIMER
        [15]   // OVERFLOW TANK DRAIN PUMP ON-DELAY
        [36]   // PANELVIEW RTC HOURLY UPDATE FROM PLC TIMER
        [16]   // OVERFLOW TANK DRAIN PUMP OFF-DELAY
        [25]   // CHEM #1 CONDUCTIVITY AT SETPOINT DELAY
        [37]   // PANELVIEW RTC HOURLY UPDATE SIGNAL TIMER
        [3]   // FORCE STEP TIMER ACC-PRE DELAY
        [17]   // OVERFLOW TANK HIGH LEVEL
        [11]   // SUPPLY TEMPERATURE AT SETPOINT DELAY
        [47].PRE   // CHEM #2 PUMP INJECTION TIME
        [18]   // PROCESS HEARTBEAT MISSING
        [48].PRE   // CHEM #2 MIX TIME
        [20]   // POWER ON DWELL DONE
        [12]   // RETURN TEMPERATURE AT SETPOINT DELAY
        [30]   // CHEM #2 CONDUCTIVITY AT SETPOINT DELAY
        [2]   // SEPARATOR TANK LOW LEVEL ALARM DELAY
        [8]   // SEPARATOR LOW LEVEL DELAY
        [4]   // SUPPLY PUMP DELAY
        [38]   // UPDATE CLOCK BUTTON VISIBLITY
   Timer_Chem1_Pump : TIMER[7] := ([0].PRE := 1000, [1].PRE := 15000, [2].PRE := 45000, [3].PRE := 5000, [4].PRE := 15000, [5].PRE := 1000, [5].ACC := 1000);   // CHEM #1 CONTROL TIMERS
        [3]   // CHEM #1 PUMP BURST ON
        [0]   // CHEM #1 PUMP DELAY ON
        [4]   // CHEM #1 PUMP BURST OFF
        [1]   // CHEM #1 INJECTION TIME
        [5]   // CHEM #1 BLOCK VALVE OFF DELAY
        [2]   // CHEM #1 MIX TIME
   Timer_Chem2_Pump : TIMER[7] := ([0].PRE := 1000, [1].PRE := 10000, [2].PRE := 50000, [3].PRE := 3000, [4].PRE := 17000, [5].PRE := 1000, [5].ACC := 1000);   // CHEM #2 CONTROL TIMERS
        [3]   // CHEM #2 PUMP BURST ON
        [0]   // CHEM #2 PUMP DELAY ON
        [4]   // CHEM #2 PUMP BURST OFF
        [5]   // CHEM #2 BLOCK VALVE OFF DELAY
        [1]   // CHEM #2 INJECTION TIME
        [2]   // CHEM #2 MIX TIME
   User_Security_Name_Display : STRING := '2';
   Utility_Button : DINT[5];   // PANELVIEW UTILITY BUTTONS
        [0].5   // PANELVIEW UTILITY BUTTON SPARE
        [0].1   // PANELVIEW UTILITY BUTTON SEPARATOR TANK DRAIN
        [0].4   // PANELVIEW UTILITY BUTTON AWFI FILL
        [0]   // SEPERATOR UTILITY BUTTONS
        [0].0   // PANELVIEW UTILITY BUTTON PW WATER FILL
        [0].2   // PANELVIEW UTILITY BUTTON CHEM #1 PUMP
        [0].3   // PANELVIEW UTILITY BUTTON CHEM #2 PUMP
   Utility_Button_Ons : DINT[5];   // PANELVIEW UTILITY BUTTON ONE SHOTS
        [0].1   // PANELVIEW UTILITY BUTTON ONE SHOT
        [0].3   // PANELVIEW UTILITY BUTTON ONE SHOT
        [0].4   // PANELVIEW UTILITY BUTTON ONE SHOT
        [0].5   // PANELVIEW UTILITY BUTTON ONE SHOT
        [0].0   // PANELVIEW UTILITY BUTTON ONE SHOT
        [0].2   // PANELVIEW UTILITY BUTTON ONE SHOT
   Utility_Ons : DINT[5];   // PANELVIEW UTILITY ONE SHOTS
        [0].1   // ONE SHOT
        [0].2   // ONE SHOT
        [0].0   // ONE SHOT
        [0].4   // ONE SHOT
        [0].5   // ONE SHOT
        [0].3   // ONE SHOT
   Utility_Out : DINT[5];   // PANELVIEW UTILITY OUTPUT CONTROL
        [0].4   // PANELVIEW UTILITY BUTTON AWFI FILL
        [0].5   // PANELVIEW UTILITY SPARE
        [0].1   // PANELVIEW UTILITY BUTTON SEPARATOR TANK DRAIN
        [0].0   // PANELVIEW UTILITY BUTTON PW WATER FILL
        [0].2   // PANELVIEW UTILITY BUTTON CHEM #1 PUMP
        [0].3   // PANELVIEW UTILITY BUTTON CHEM #2 PUMP
   Utility_Timer : TIMER[4] := ([0].PRE := 20000, [1].PRE := 20000, [2].PRE := 20000, [3].PRE := 20000);   // PANELVIEW UTILITY TIMERS
        [1]   // PANELVIEW UTILITY CHEM #2 PUMP DELAY OFF
        [0]   // PANELVIEW UTILITY CHEM #1 PUMP DELAY OFF
END_VAR
